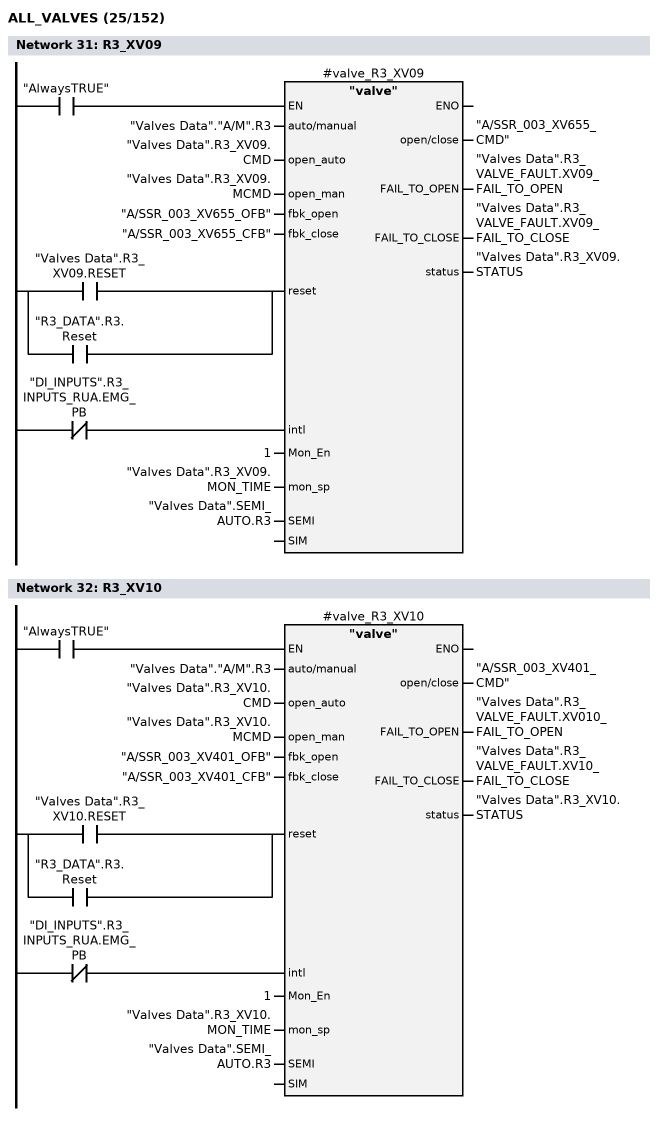
   RUNG wire#powerrail
      Contact( "AlwaysTRUE" )
      #valve_R3_XV09(reset := wire#w1, intl := wire#w2, "auto/manual" := "Valves Data"."A/M".R3, open_auto := "Valves Data".R3_XV09.CMD, open_man := "Valves Data".R3_XV09.MCMD, fbk_open := "A/SSR_003_XV655_OFB", fbk_close := "A/SSR_003_XV655_CFB", Mon_En := 1, mon_sp := "Valves Data".R3_XV09.MON_TIME, SEMI := "Valves Data".SEMI_AUTO.R3, SIM :=, "open/close" => "A/SSR_003_XV655_CMD", FAIL_TO_OPEN => "Valves Data".R3_VALVE_FAULT.XV09_FAIL_TO_OPEN, FAIL_TO_CLOSE => "Valves Data".R3_VALVE_FAULT.XV09_FAIL_TO_CLOSE, status => "Valves Data".R3_XV09.STATUS)
   END_RUNG
   RUNG wire#powerrail
      Contact( "Valves Data".R3_XV09.RESET )
   END_RUNG wire#w1
   RUNG wire#powerrail
      Contact( "R3_DATA".R3.Reset )
   END_RUNG wire#w1
   RUNG wire#powerrail
      I_Contact( "DI_INPUTS".R3_INPUTS_RUA.EMG_PB )
   END_RUNG wire#w2
   // the same network as SCL:
   IF "AlwaysTRUE" THEN
       #valve_R3_XV09("auto/manual" := "Valves Data"."A/M".R3,   // "valve"
                      open_auto := "Valves Data".R3_XV09.CMD,
                      open_man := "Valves Data".R3_XV09.MCMD,
                      fbk_open := "A/SSR_003_XV655_OFB",
                      fbk_close := "A/SSR_003_XV655_CFB",
                      reset := "Valves Data".R3_XV09.RESET OR "R3_DATA".R3.Reset,
                      intl := NOT "DI_INPUTS".R3_INPUTS_RUA.EMG_PB,
                      Mon_En := 1,
                      mon_sp := "Valves Data".R3_XV09.MON_TIME,
                      SEMI := "Valves Data".SEMI_AUTO.R3,
                      "open/close" => "A/SSR_003_XV655_CMD",
                      FAIL_TO_OPEN => "Valves Data".R3_VALVE_FAULT.XV09_FAIL_TO_OPEN,
                      FAIL_TO_CLOSE => "Valves Data".R3_VALVE_FAULT.XV09_FAIL_TO_CLOSE,
                      status => "Valves Data".R3_XV09.STATUS);
   END_IF;
END_REGION

REGION Network 32: R3_XV10
   RUNG wire#powerrail
      Contact( "AlwaysTRUE" )
      #valve_R3_XV10(reset := wire#w1, intl := wire#w2, "auto/manual" := "Valves Data"."A/M".R3, open_auto := "Valves Data".R3_XV10.CMD, open_man := "Valves Data".R3_XV10.MCMD, fbk_open := "A/SSR_003_XV401_OFB", fbk_close := "A/SSR_003_XV401_CFB", Mon_En := 1, mon_sp := "Valves Data".R3_XV10.MON_TIME, SEMI := "Valves Data".SEMI_AUTO.R3, SIM :=, "open/close" => "A/SSR_003_XV401_CMD", FAIL_TO_OPEN => "Valves Data".R3_VALVE_FAULT.XV010_FAIL_TO_OPEN, FAIL_TO_CLOSE => "Valves Data".R3_VALVE_FAULT.XV10_FAIL_TO_CLOSE, status => "Valves Data".R3_XV10.STATUS)
   END_RUNG
   RUNG wire#powerrail
      Contact( "Valves Data".R3_XV10.RESET )
   END_RUNG wire#w1
   RUNG wire#powerrail
      Contact( "R3_DATA".R3.Reset )
   END_RUNG wire#w1
   RUNG wire#powerrail
      I_Contact( "DI_INPUTS".R3_INPUTS_RUA.EMG_PB )
   END_RUNG wire#w2
   // the same network as SCL:
   IF "AlwaysTRUE" THEN
       #valve_R3_XV10("auto/manual" := "Valves Data"."A/M".R3,   // "valve"
                      open_auto := "Valves Data".R3_XV10.CMD,
                      open_man := "Valves Data".R3_XV10.MCMD,
                      fbk_open := "A/SSR_003_XV401_OFB",
                      fbk_close := "A/SSR_003_XV401_CFB",
                      reset := "Valves Data".R3_XV10.RESET OR "R3_DATA".R3.Reset,
                      intl := NOT "DI_INPUTS".R3_INPUTS_RUA.EMG_PB,
                      Mon_En := 1,
                      mon_sp := "Valves Data".R3_XV10.MON_TIME,
                      SEMI := "Valves Data".SEMI_AUTO.R3,
                      "open/close" => "A/SSR_003_XV401_CMD",
                      FAIL_TO_OPEN => "Valves Data".R3_VALVE_FAULT.XV010_FAIL_TO_OPEN,
                      FAIL_TO_CLOSE => "Valves Data".R3_VALVE_FAULT.XV10_FAIL_TO_CLOSE,
                      status => "Valves Data".R3_XV10.STATUS);
   END_IF;
END_REGION

REGION Network 33: ****REACTOR_04****
END_REGION

REGION Network 34: R4_XV01
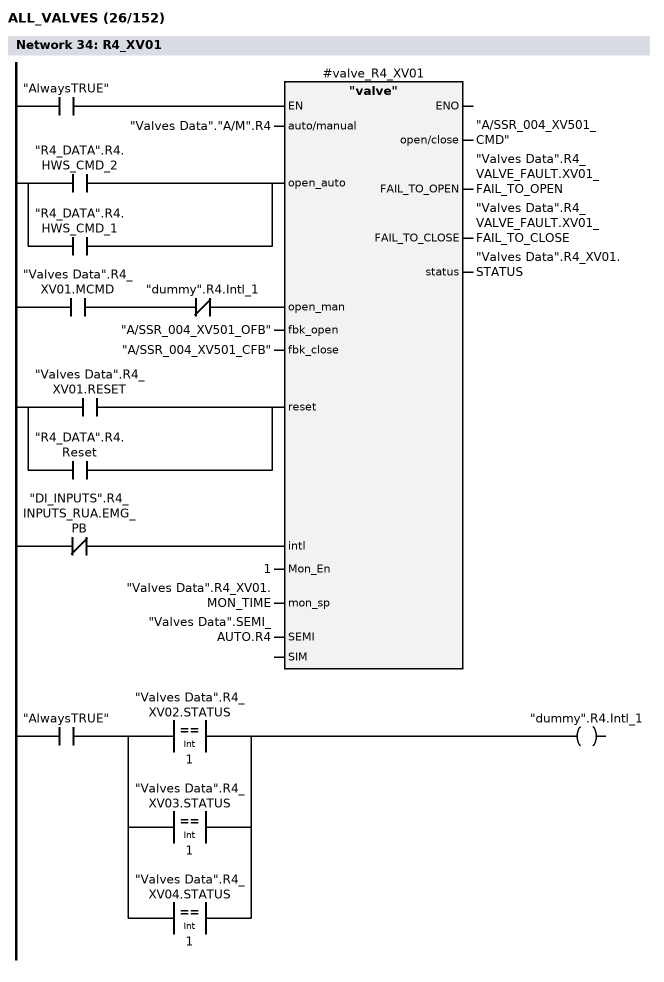
   RUNG wire#powerrail
      Contact( "AlwaysTRUE" )
      #valve_R4_XV01(open_auto := wire#w1, open_man := wire#w2, reset := wire#w3, intl := wire#w4, "auto/manual" := "Valves Data"."A/M".R4, fbk_open := "A/SSR_004_XV501_OFB", fbk_close := "A/SSR_004_XV501_CFB", Mon_En := 1, mon_sp := "Valves Data".R4_XV01.MON_TIME, SEMI := "Valves Data".SEMI_AUTO.R4, SIM :=, "open/close" => "A/SSR_004_XV501_CMD", FAIL_TO_OPEN => "Valves Data".R4_VALVE_FAULT.XV01_FAIL_TO_OPEN, FAIL_TO_CLOSE => "Valves Data".R4_VALVE_FAULT.XV01_FAIL_TO_CLOSE, status => "Valves Data".R4_XV01.STATUS)
   END_RUNG
   RUNG wire#powerrail
      Contact( "R4_DATA".R4.HWS_CMD_2 )
   END_RUNG wire#w1
   RUNG wire#powerrail
      Contact( "R4_DATA".R4.HWS_CMD_1 )
   END_RUNG wire#w1
   RUNG wire#powerrail
      Contact( "Valves Data".R4_XV01.MCMD )
      I_Contact( "dummy".R4.Intl_1 )
   END_RUNG wire#w2
   RUNG wire#powerrail
      Contact( "Valves Data".R4_XV01.RESET )
   END_RUNG wire#w3
   RUNG wire#powerrail
      Contact( "R4_DATA".R4.Reset )
   END_RUNG wire#w3
   RUNG wire#powerrail
      I_Contact( "DI_INPUTS".R4_INPUTS_RUA.EMG_PB )
   END_RUNG wire#w4
   RUNG wire#powerrail
      Contact( "AlwaysTRUE" )
      wire#w5
      { S7_Templates := "SrcType := Int" } EQ_Contact(in1 := "Valves Data".R4_XV02.STATUS, in2 := 1)
      wire#w6
      Coil( "dummy".R4.Intl_1 )
   END_RUNG
   RUNG wire#w5
      { S7_Templates := "SrcType := Int" } EQ_Contact(in1 := "Valves Data".R4_XV03.STATUS, in2 := 1)
   END_RUNG wire#w6
   RUNG wire#w5
      { S7_Templates := "SrcType := Int" } EQ_Contact(in1 := "Valves Data".R4_XV04.STATUS, in2 := 1)
   END_RUNG wire#w6
   // the same network as SCL:
   IF "AlwaysTRUE" THEN
       #valve_R4_XV01("auto/manual" := "Valves Data"."A/M".R4,   // "valve"
                      open_auto := "R4_DATA".R4.HWS_CMD_2 OR "R4_DATA".R4.HWS_CMD_1,
                      open_man := "Valves Data".R4_XV01.MCMD AND NOT "dummy".R4.Intl_1,
                      fbk_open := "A/SSR_004_XV501_OFB",
                      fbk_close := "A/SSR_004_XV501_CFB",
                      reset := "Valves Data".R4_XV01.RESET OR "R4_DATA".R4.Reset,
                      intl := NOT "DI_INPUTS".R4_INPUTS_RUA.EMG_PB,
                      Mon_En := 1,
                      mon_sp := "Valves Data".R4_XV01.MON_TIME,
                      SEMI := "Valves Data".SEMI_AUTO.R4,
                      "open/close" => "A/SSR_004_XV501_CMD",
                      FAIL_TO_OPEN => "Valves Data".R4_VALVE_FAULT.XV01_FAIL_TO_OPEN,
                      FAIL_TO_CLOSE => "Valves Data".R4_VALVE_FAULT.XV01_FAIL_TO_CLOSE,
                      status => "Valves Data".R4_XV01.STATUS);
   END_IF;
   "dummy".R4.Intl_1 := "AlwaysTRUE" AND (("Valves Data".R4_XV02.STATUS = 1) OR ("Valves Data".R4_XV03.STATUS = 1) OR ("Valves Data".R4_XV04.STATUS = 1));
END_REGION

REGION Network 35: R4_XV02
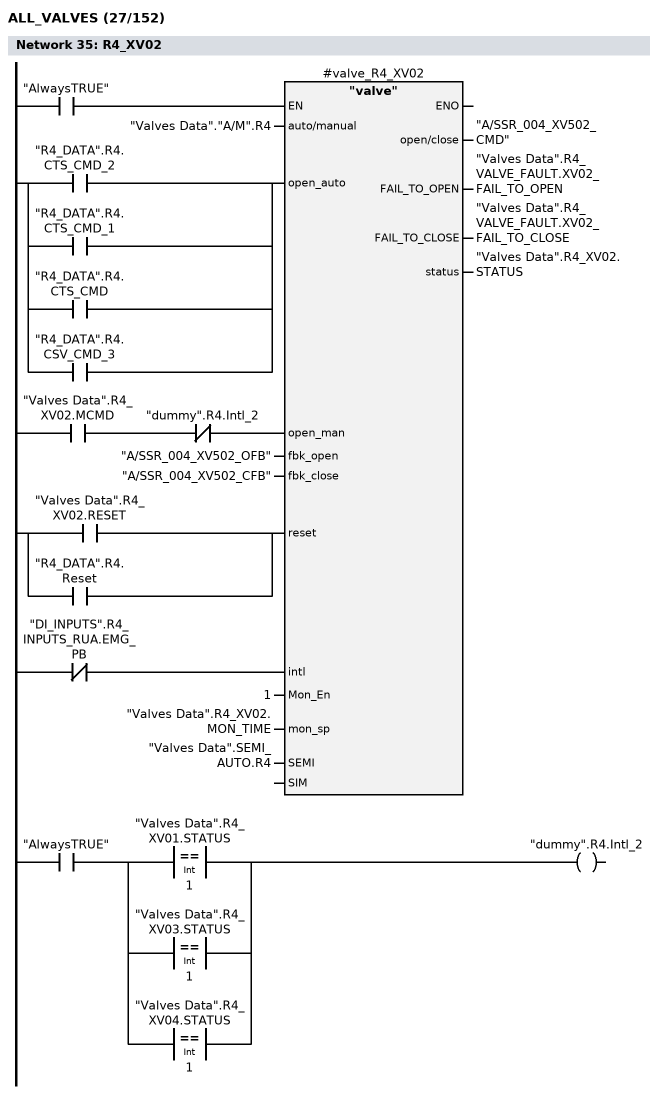
   RUNG wire#powerrail
      Contact( "AlwaysTRUE" )
      #valve_R4_XV02(open_auto := wire#w1, open_man := wire#w2, reset := wire#w3, intl := wire#w4, "auto/manual" := "Valves Data"."A/M".R4, fbk_open := "A/SSR_004_XV502_OFB", fbk_close := "A/SSR_004_XV502_CFB", Mon_En := 1, mon_sp := "Valves Data".R4_XV02.MON_TIME, SEMI := "Valves Data".SEMI_AUTO.R4, SIM :=, "open/close" => "A/SSR_004_XV502_CMD", FAIL_TO_OPEN => "Valves Data".R4_VALVE_FAULT.XV02_FAIL_TO_OPEN, FAIL_TO_CLOSE => "Valves Data".R4_VALVE_FAULT.XV02_FAIL_TO_CLOSE, status => "Valves Data".R4_XV02.STATUS)
   END_RUNG
   RUNG wire#powerrail
      Contact( "R4_DATA".R4.CTS_CMD_2 )
   END_RUNG wire#w1
   RUNG wire#powerrail
      Contact( "R4_DATA".R4.CTS_CMD_1 )
   END_RUNG wire#w1
   RUNG wire#powerrail
      Contact( "R4_DATA".R4.CTS_CMD )
   END_RUNG wire#w1
   RUNG wire#powerrail
      Contact( "R4_DATA".R4.CSV_CMD_3 )
   END_RUNG wire#w1
   RUNG wire#powerrail
      Contact( "Valves Data".R4_XV02.MCMD )
      I_Contact( "dummy".R4.Intl_2 )
   END_RUNG wire#w2
   RUNG wire#powerrail
      Contact( "Valves Data".R4_XV02.RESET )
   END_RUNG wire#w3
   RUNG wire#powerrail
      Contact( "R4_DATA".R4.Reset )
   END_RUNG wire#w3
   RUNG wire#powerrail
      I_Contact( "DI_INPUTS".R4_INPUTS_RUA.EMG_PB )
   END_RUNG wire#w4
   RUNG wire#powerrail
      Contact( "AlwaysTRUE" )
      wire#w5
      { S7_Templates := "SrcType := Int" } EQ_Contact(in1 := "Valves Data".R4_XV01.STATUS, in2 := 1)
      wire#w6
      Coil( "dummy".R4.Intl_2 )
   END_RUNG
   RUNG wire#w5
      { S7_Templates := "SrcType := Int" } EQ_Contact(in1 := "Valves Data".R4_XV03.STATUS, in2 := 1)
   END_RUNG wire#w6
   RUNG wire#w5
      { S7_Templates := "SrcType := Int" } EQ_Contact(in1 := "Valves Data".R4_XV04.STATUS, in2 := 1)
   END_RUNG wire#w6
   // the same network as SCL:
   IF "AlwaysTRUE" THEN
       #valve_R4_XV02("auto/manual" := "Valves Data"."A/M".R4,   // "valve"
                      open_auto := "R4_DATA".R4.CTS_CMD_2 OR "R4_DATA".R4.CTS_CMD_1 OR "R4_DATA".R4.CTS_CMD OR "R4_DATA".R4.CSV_CMD_3,
                      open_man := "Valves Data".R4_XV02.MCMD AND NOT "dummy".R4.Intl_2,
                      fbk_open := "A/SSR_004_XV502_OFB",
                      fbk_close := "A/SSR_004_XV502_CFB",
                      reset := "Valves Data".R4_XV02.RESET OR "R4_DATA".R4.Reset,
                      intl := NOT "DI_INPUTS".R4_INPUTS_RUA.EMG_PB,
                      Mon_En := 1,
                      mon_sp := "Valves Data".R4_XV02.MON_TIME,
                      SEMI := "Valves Data".SEMI_AUTO.R4,
                      "open/close" => "A/SSR_004_XV502_CMD",
                      FAIL_TO_OPEN => "Valves Data".R4_VALVE_FAULT.XV02_FAIL_TO_OPEN,
                      FAIL_TO_CLOSE => "Valves Data".R4_VALVE_FAULT.XV02_FAIL_TO_CLOSE,
                      status => "Valves Data".R4_XV02.STATUS);
   END_IF;
   "dummy".R4.Intl_2 := "AlwaysTRUE" AND (("Valves Data".R4_XV01.STATUS = 1) OR ("Valves Data".R4_XV03.STATUS = 1) OR ("Valves Data".R4_XV04.STATUS = 1));
END_REGION

REGION Network 36: R4_XV03
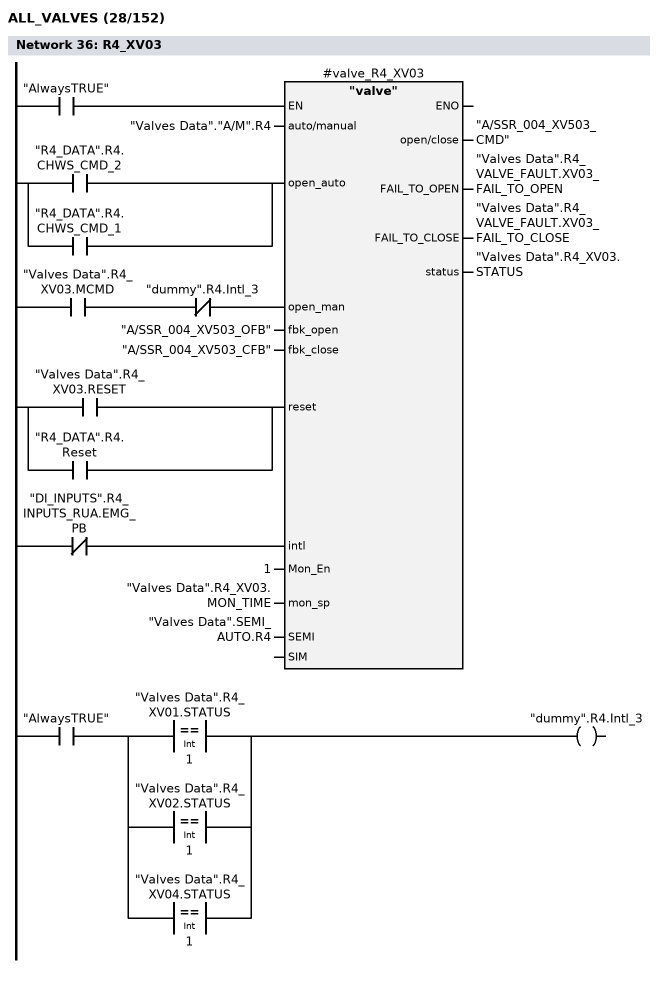
   RUNG wire#powerrail
      Contact( "AlwaysTRUE" )
      #valve_R4_XV03(open_auto := wire#w1, open_man := wire#w2, reset := wire#w3, intl := wire#w4, "auto/manual" := "Valves Data"."A/M".R4, fbk_open := "A/SSR_004_XV503_OFB", fbk_close := "A/SSR_004_XV503_CFB", Mon_En := 1, mon_sp := "Valves Data".R4_XV03.MON_TIME, SEMI := "Valves Data".SEMI_AUTO.R4, SIM :=, "open/close" => "A/SSR_004_XV503_CMD", FAIL_TO_OPEN => "Valves Data".R4_VALVE_FAULT.XV03_FAIL_TO_OPEN, FAIL_TO_CLOSE => "Valves Data".R4_VALVE_FAULT.XV03_FAIL_TO_CLOSE, status => "Valves Data".R4_XV03.STATUS)
   END_RUNG
   RUNG wire#powerrail
      Contact( "R4_DATA".R4.CHWS_CMD_2 )
   END_RUNG wire#w1
   RUNG wire#powerrail
      Contact( "R4_DATA".R4.CHWS_CMD_1 )
   END_RUNG wire#w1
   RUNG wire#powerrail
      Contact( "Valves Data".R4_XV03.MCMD )
      I_Contact( "dummy".R4.Intl_3 )
   END_RUNG wire#w2
   RUNG wire#powerrail
      Contact( "Valves Data".R4_XV03.RESET )
   END_RUNG wire#w3
   RUNG wire#powerrail
      Contact( "R4_DATA".R4.Reset )
   END_RUNG wire#w3
   RUNG wire#powerrail
      I_Contact( "DI_INPUTS".R4_INPUTS_RUA.EMG_PB )
   END_RUNG wire#w4
   RUNG wire#powerrail
      Contact( "AlwaysTRUE" )
      wire#w5
      { S7_Templates := "SrcType := Int" } EQ_Contact(in1 := "Valves Data".R4_XV01.STATUS, in2 := 1)
      wire#w6
      Coil( "dummy".R4.Intl_3 )
   END_RUNG
   RUNG wire#w5
      { S7_Templates := "SrcType := Int" } EQ_Contact(in1 := "Valves Data".R4_XV02.STATUS, in2 := 1)
   END_RUNG wire#w6
   RUNG wire#w5
      { S7_Templates := "SrcType := Int" } EQ_Contact(in1 := "Valves Data".R4_XV04.STATUS, in2 := 1)
   END_RUNG wire#w6
   // the same network as SCL:
   IF "AlwaysTRUE" THEN
       #valve_R4_XV03("auto/manual" := "Valves Data"."A/M".R4,   // "valve"
                      open_auto := "R4_DATA".R4.CHWS_CMD_2 OR "R4_DATA".R4.CHWS_CMD_1,
                      open_man := "Valves Data".R4_XV03.MCMD AND NOT "dummy".R4.Intl_3,
                      fbk_open := "A/SSR_004_XV503_OFB",
                      fbk_close := "A/SSR_004_XV503_CFB",
                      reset := "Valves Data".R4_XV03.RESET OR "R4_DATA".R4.Reset,
                      intl := NOT "DI_INPUTS".R4_INPUTS_RUA.EMG_PB,
                      Mon_En := 1,
                      mon_sp := "Valves Data".R4_XV03.MON_TIME,
                      SEMI := "Valves Data".SEMI_AUTO.R4,
                      "open/close" => "A/SSR_004_XV503_CMD",
                      FAIL_TO_OPEN => "Valves Data".R4_VALVE_FAULT.XV03_FAIL_TO_OPEN,
                      FAIL_TO_CLOSE => "Valves Data".R4_VALVE_FAULT.XV03_FAIL_TO_CLOSE,
                      status => "Valves Data".R4_XV03.STATUS);
   END_IF;
   "dummy".R4.Intl_3 := "AlwaysTRUE" AND (("Valves Data".R4_XV01.STATUS = 1) OR ("Valves Data".R4_XV02.STATUS = 1) OR ("Valves Data".R4_XV04.STATUS = 1));
END_REGION

REGION Network 37: R4_XV04
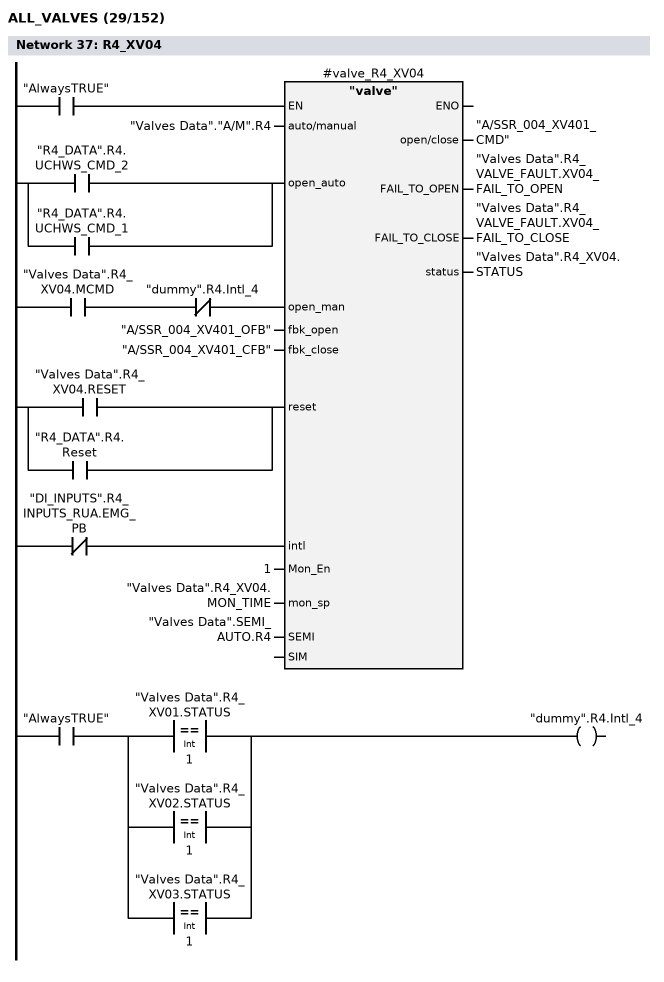
   RUNG wire#powerrail
      Contact( "AlwaysTRUE" )
      #valve_R4_XV04(open_auto := wire#w1, open_man := wire#w2, reset := wire#w3, intl := wire#w4, "auto/manual" := "Valves Data"."A/M".R4, fbk_open := "A/SSR_004_XV401_OFB", fbk_close := "A/SSR_004_XV401_CFB", Mon_En := 1, mon_sp := "Valves Data".R4_XV04.MON_TIME, SEMI := "Valves Data".SEMI_AUTO.R4, SIM :=, "open/close" => "A/SSR_004_XV401_CMD", FAIL_TO_OPEN => "Valves Data".R4_VALVE_FAULT.XV04_FAIL_TO_OPEN, FAIL_TO_CLOSE => "Valves Data".R4_VALVE_FAULT.XV04_FAIL_TO_CLOSE, status => "Valves Data".R4_XV04.STATUS)
   END_RUNG
   RUNG wire#powerrail
      Contact( "R4_DATA".R4.UCHWS_CMD_2 )
   END_RUNG wire#w1
   RUNG wire#powerrail
      Contact( "R4_DATA".R4.UCHWS_CMD_1 )
   END_RUNG wire#w1
   RUNG wire#powerrail
      Contact( "Valves Data".R4_XV04.MCMD )
      I_Contact( "dummy".R4.Intl_4 )
   END_RUNG wire#w2
   RUNG wire#powerrail
      Contact( "Valves Data".R4_XV04.RESET )
   END_RUNG wire#w3
   RUNG wire#powerrail
      Contact( "R4_DATA".R4.Reset )
   END_RUNG wire#w3
   RUNG wire#powerrail
      I_Contact( "DI_INPUTS".R4_INPUTS_RUA.EMG_PB )
   END_RUNG wire#w4
   RUNG wire#powerrail
      Contact( "AlwaysTRUE" )
      wire#w5
      { S7_Templates := "SrcType := Int" } EQ_Contact(in1 := "Valves Data".R4_XV01.STATUS, in2 := 1)
      wire#w6
      Coil( "dummy".R4.Intl_4 )
   END_RUNG
   RUNG wire#w5
      { S7_Templates := "SrcType := Int" } EQ_Contact(in1 := "Valves Data".R4_XV02.STATUS, in2 := 1)
   END_RUNG wire#w6
   RUNG wire#w5
      { S7_Templates := "SrcType := Int" } EQ_Contact(in1 := "Valves Data".R4_XV03.STATUS, in2 := 1)
   END_RUNG wire#w6
   // the same network as SCL:
   IF "AlwaysTRUE" THEN
       #valve_R4_XV04("auto/manual" := "Valves Data"."A/M".R4,   // "valve"
                      open_auto := "R4_DATA".R4.UCHWS_CMD_2 OR "R4_DATA".R4.UCHWS_CMD_1,
                      open_man := "Valves Data".R4_XV04.MCMD AND NOT "dummy".R4.Intl_4,
                      fbk_open := "A/SSR_004_XV401_OFB",
                      fbk_close := "A/SSR_004_XV401_CFB",
                      reset := "Valves Data".R4_XV04.RESET OR "R4_DATA".R4.Reset,
                      intl := NOT "DI_INPUTS".R4_INPUTS_RUA.EMG_PB,
                      Mon_En := 1,
                      mon_sp := "Valves Data".R4_XV04.MON_TIME,
                      SEMI := "Valves Data".SEMI_AUTO.R4,
                      "open/close" => "A/SSR_004_XV401_CMD",
                      FAIL_TO_OPEN => "Valves Data".R4_VALVE_FAULT.XV04_FAIL_TO_OPEN,
                      FAIL_TO_CLOSE => "Valves Data".R4_VALVE_FAULT.XV04_FAIL_TO_CLOSE,
                      status => "Valves Data".R4_XV04.STATUS);
   END_IF;
   "dummy".R4.Intl_4 := "AlwaysTRUE" AND (("Valves Data".R4_XV01.STATUS = 1) OR ("Valves Data".R4_XV02.STATUS = 1) OR ("Valves Data".R4_XV03.STATUS = 1));
END_REGION

REGION Network 38: R4_XV05
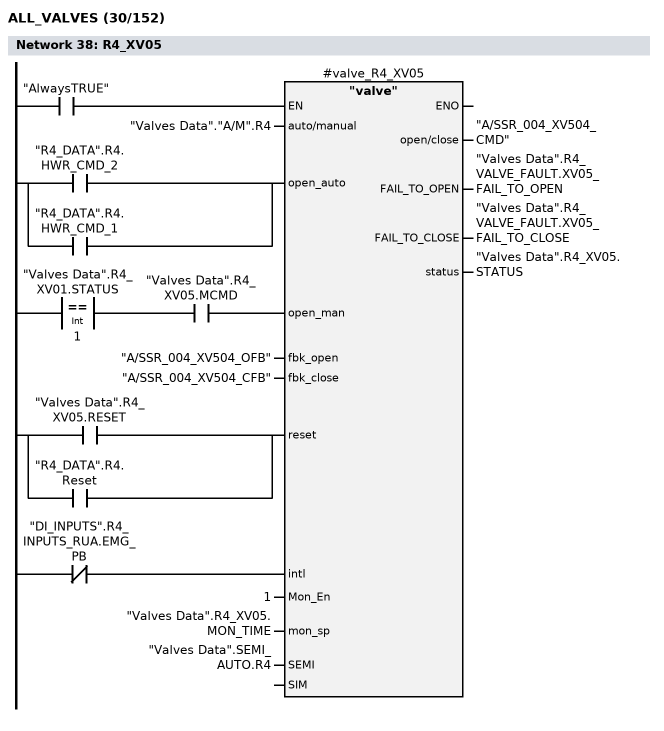
   RUNG wire#powerrail
      Contact( "AlwaysTRUE" )
      #valve_R4_XV05(open_auto := wire#w1, open_man := wire#w2, reset := wire#w3, intl := wire#w4, "auto/manual" := "Valves Data"."A/M".R4, fbk_open := "A/SSR_004_XV504_OFB", fbk_close := "A/SSR_004_XV504_CFB", Mon_En := 1, mon_sp := "Valves Data".R4_XV05.MON_TIME, SEMI := "Valves Data".SEMI_AUTO.R4, SIM :=, "open/close" => "A/SSR_004_XV504_CMD", FAIL_TO_OPEN => "Valves Data".R4_VALVE_FAULT.XV05_FAIL_TO_OPEN, FAIL_TO_CLOSE => "Valves Data".R4_VALVE_FAULT.XV05_FAIL_TO_CLOSE, status => "Valves Data".R4_XV05.STATUS)
   END_RUNG
   RUNG wire#powerrail
      Contact( "R4_DATA".R4.HWR_CMD_2 )
   END_RUNG wire#w1
   RUNG wire#powerrail
      Contact( "R4_DATA".R4.HWR_CMD_1 )
   END_RUNG wire#w1
   RUNG wire#powerrail
      { S7_Templates := "SrcType := Int" } EQ_Contact(in1 := "Valves Data".R4_XV01.STATUS, in2 := 1)
      Contact( "Valves Data".R4_XV05.MCMD )
   END_RUNG wire#w2
   RUNG wire#powerrail
      Contact( "Valves Data".R4_XV05.RESET )
   END_RUNG wire#w3
   RUNG wire#powerrail
      Contact( "R4_DATA".R4.Reset )
   END_RUNG wire#w3
   RUNG wire#powerrail
      I_Contact( "DI_INPUTS".R4_INPUTS_RUA.EMG_PB )
   END_RUNG wire#w4
   // the same network as SCL:
   IF "AlwaysTRUE" THEN
       #valve_R4_XV05("auto/manual" := "Valves Data"."A/M".R4,   // "valve"
                      open_auto := "R4_DATA".R4.HWR_CMD_2 OR "R4_DATA".R4.HWR_CMD_1,
                      open_man := ("Valves Data".R4_XV01.STATUS = 1) AND "Valves Data".R4_XV05.MCMD,
                      fbk_open := "A/SSR_004_XV504_OFB",
                      fbk_close := "A/SSR_004_XV504_CFB",
                      reset := "Valves Data".R4_XV05.RESET OR "R4_DATA".R4.Reset,
                      intl := NOT "DI_INPUTS".R4_INPUTS_RUA.EMG_PB,
                      Mon_En := 1,
                      mon_sp := "Valves Data".R4_XV05.MON_TIME,
                      SEMI := "Valves Data".SEMI_AUTO.R4,
                      "open/close" => "A/SSR_004_XV504_CMD",
                      FAIL_TO_OPEN => "Valves Data".R4_VALVE_FAULT.XV05_FAIL_TO_OPEN,
                      FAIL_TO_CLOSE => "Valves Data".R4_VALVE_FAULT.XV05_FAIL_TO_CLOSE,
                      status => "Valves Data".R4_XV05.STATUS);
   END_IF;
END_REGION

REGION Network 39: R4_XV06
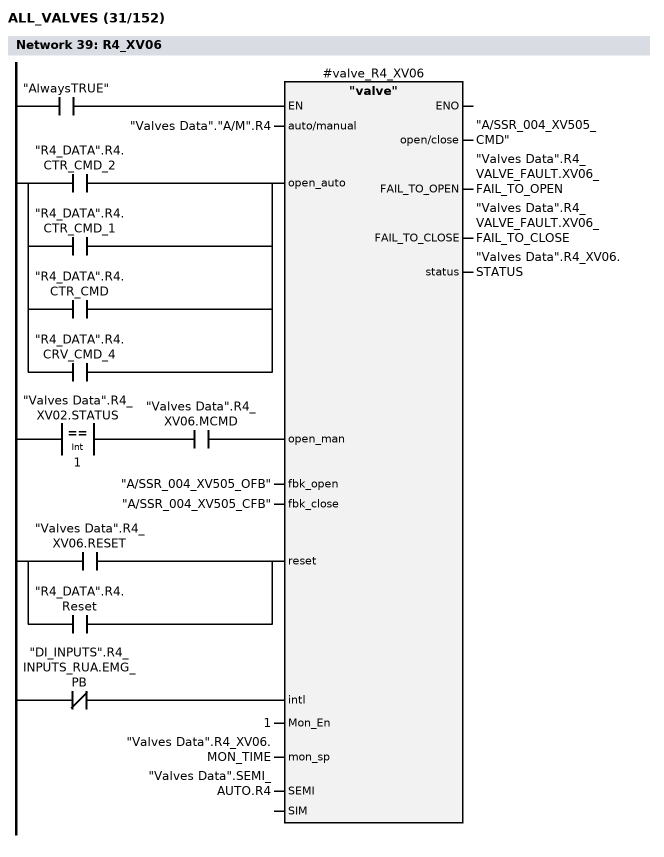
   RUNG wire#powerrail
      Contact( "AlwaysTRUE" )
      #valve_R4_XV06(open_auto := wire#w1, open_man := wire#w2, reset := wire#w3, intl := wire#w4, "auto/manual" := "Valves Data"."A/M".R4, fbk_open := "A/SSR_004_XV505_OFB", fbk_close := "A/SSR_004_XV505_CFB", Mon_En := 1, mon_sp := "Valves Data".R4_XV06.MON_TIME, SEMI := "Valves Data".SEMI_AUTO.R4, SIM :=, "open/close" => "A/SSR_004_XV505_CMD", FAIL_TO_OPEN => "Valves Data".R4_VALVE_FAULT.XV06_FAIL_TO_OPEN, FAIL_TO_CLOSE => "Valves Data".R4_VALVE_FAULT.XV06_FAIL_TO_CLOSE, status => "Valves Data".R4_XV06.STATUS)
   END_RUNG
   RUNG wire#powerrail
      Contact( "R4_DATA".R4.CTR_CMD_2 )
   END_RUNG wire#w1
   RUNG wire#powerrail
      Contact( "R4_DATA".R4.CTR_CMD_1 )
   END_RUNG wire#w1
   RUNG wire#powerrail
      Contact( "R4_DATA".R4.CTR_CMD )
   END_RUNG wire#w1
   RUNG wire#powerrail
      Contact( "R4_DATA".R4.CRV_CMD_4 )
   END_RUNG wire#w1
   RUNG wire#powerrail
      { S7_Templates := "SrcType := Int" } EQ_Contact(in1 := "Valves Data".R4_XV02.STATUS, in2 := 1)
      Contact( "Valves Data".R4_XV06.MCMD )
   END_RUNG wire#w2
   RUNG wire#powerrail
      Contact( "Valves Data".R4_XV06.RESET )
   END_RUNG wire#w3
   RUNG wire#powerrail
      Contact( "R4_DATA".R4.Reset )
   END_RUNG wire#w3
   RUNG wire#powerrail
      I_Contact( "DI_INPUTS".R4_INPUTS_RUA.EMG_PB )
   END_RUNG wire#w4
   // the same network as SCL:
   IF "AlwaysTRUE" THEN
       #valve_R4_XV06("auto/manual" := "Valves Data"."A/M".R4,   // "valve"
                      open_auto := "R4_DATA".R4.CTR_CMD_2 OR "R4_DATA".R4.CTR_CMD_1 OR "R4_DATA".R4.CTR_CMD OR "R4_DATA".R4.CRV_CMD_4,
                      open_man := ("Valves Data".R4_XV02.STATUS = 1) AND "Valves Data".R4_XV06.MCMD,
                      fbk_open := "A/SSR_004_XV505_OFB",
                      fbk_close := "A/SSR_004_XV505_CFB",
                      reset := "Valves Data".R4_XV06.RESET OR "R4_DATA".R4.Reset,
                      intl := NOT "DI_INPUTS".R4_INPUTS_RUA.EMG_PB,
                      Mon_En := 1,
                      mon_sp := "Valves Data".R4_XV06.MON_TIME,
                      SEMI := "Valves Data".SEMI_AUTO.R4,
                      "open/close" => "A/SSR_004_XV505_CMD",
                      FAIL_TO_OPEN => "Valves Data".R4_VALVE_FAULT.XV06_FAIL_TO_OPEN,
                      FAIL_TO_CLOSE => "Valves Data".R4_VALVE_FAULT.XV06_FAIL_TO_CLOSE,
                      status => "Valves Data".R4_XV06.STATUS);
   END_IF;
END_REGION

REGION Network 40: R4_XV07
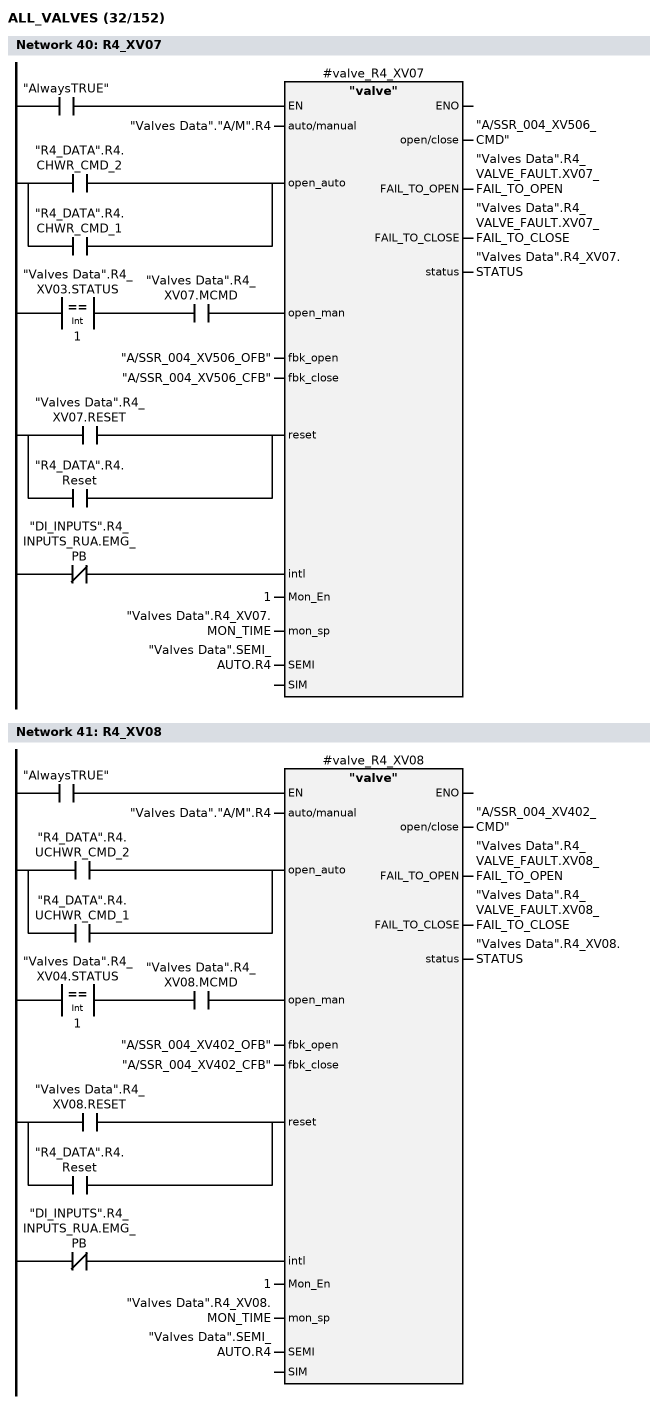
   RUNG wire#powerrail
      Contact( "AlwaysTRUE" )
      #valve_R4_XV07(open_auto := wire#w1, open_man := wire#w2, reset := wire#w3, intl := wire#w4, "auto/manual" := "Valves Data"."A/M".R4, fbk_open := "A/SSR_004_XV506_OFB", fbk_close := "A/SSR_004_XV506_CFB", Mon_En := 1, mon_sp := "Valves Data".R4_XV07.MON_TIME, SEMI := "Valves Data".SEMI_AUTO.R4, SIM :=, "open/close" => "A/SSR_004_XV506_CMD", FAIL_TO_OPEN => "Valves Data".R4_VALVE_FAULT.XV07_FAIL_TO_OPEN, FAIL_TO_CLOSE => "Valves Data".R4_VALVE_FAULT.XV07_FAIL_TO_CLOSE, status => "Valves Data".R4_XV07.STATUS)
   END_RUNG
   RUNG wire#powerrail
      Contact( "R4_DATA".R4.CHWR_CMD_2 )
   END_RUNG wire#w1
   RUNG wire#powerrail
      Contact( "R4_DATA".R4.CHWR_CMD_1 )
   END_RUNG wire#w1
   RUNG wire#powerrail
      { S7_Templates := "SrcType := Int" } EQ_Contact(in1 := "Valves Data".R4_XV03.STATUS, in2 := 1)
      Contact( "Valves Data".R4_XV07.MCMD )
   END_RUNG wire#w2
   RUNG wire#powerrail
      Contact( "Valves Data".R4_XV07.RESET )
   END_RUNG wire#w3
   RUNG wire#powerrail
      Contact( "R4_DATA".R4.Reset )
   END_RUNG wire#w3
   RUNG wire#powerrail
      I_Contact( "DI_INPUTS".R4_INPUTS_RUA.EMG_PB )
   END_RUNG wire#w4
   // the same network as SCL:
   IF "AlwaysTRUE" THEN
       #valve_R4_XV07("auto/manual" := "Valves Data"."A/M".R4,   // "valve"
                      open_auto := "R4_DATA".R4.CHWR_CMD_2 OR "R4_DATA".R4.CHWR_CMD_1,
                      open_man := ("Valves Data".R4_XV03.STATUS = 1) AND "Valves Data".R4_XV07.MCMD,
                      fbk_open := "A/SSR_004_XV506_OFB",
                      fbk_close := "A/SSR_004_XV506_CFB",
                      reset := "Valves Data".R4_XV07.RESET OR "R4_DATA".R4.Reset,
                      intl := NOT "DI_INPUTS".R4_INPUTS_RUA.EMG_PB,
                      Mon_En := 1,
                      mon_sp := "Valves Data".R4_XV07.MON_TIME,
                      SEMI := "Valves Data".SEMI_AUTO.R4,
                      "open/close" => "A/SSR_004_XV506_CMD",
                      FAIL_TO_OPEN => "Valves Data".R4_VALVE_FAULT.XV07_FAIL_TO_OPEN,
                      FAIL_TO_CLOSE => "Valves Data".R4_VALVE_FAULT.XV07_FAIL_TO_CLOSE,
                      status => "Valves Data".R4_XV07.STATUS);
   END_IF;
END_REGION

REGION Network 41: R4_XV08
   RUNG wire#powerrail
      Contact( "AlwaysTRUE" )
      #valve_R4_XV08(open_auto := wire#w1, open_man := wire#w2, reset := wire#w3, intl := wire#w4, "auto/manual" := "Valves Data"."A/M".R4, fbk_open := "A/SSR_004_XV402_OFB", fbk_close := "A/SSR_004_XV402_CFB", Mon_En := 1, mon_sp := "Valves Data".R4_XV08.MON_TIME, SEMI := "Valves Data".SEMI_AUTO.R4, SIM :=, "open/close" => "A/SSR_004_XV402_CMD", FAIL_TO_OPEN => "Valves Data".R4_VALVE_FAULT.XV08_FAIL_TO_OPEN, FAIL_TO_CLOSE => "Valves Data".R4_VALVE_FAULT.XV08_FAIL_TO_CLOSE, status => "Valves Data".R4_XV08.STATUS)
   END_RUNG
   RUNG wire#powerrail
      Contact( "R4_DATA".R4.UCHWR_CMD_2 )
   END_RUNG wire#w1
   RUNG wire#powerrail
      Contact( "R4_DATA".R4.UCHWR_CMD_1 )
   END_RUNG wire#w1
   RUNG wire#powerrail
      { S7_Templates := "SrcType := Int" } EQ_Contact(in1 := "Valves Data".R4_XV04.STATUS, in2 := 1)
      Contact( "Valves Data".R4_XV08.MCMD )
   END_RUNG wire#w2
   RUNG wire#powerrail
      Contact( "Valves Data".R4_XV08.RESET )
   END_RUNG wire#w3
   RUNG wire#powerrail
      Contact( "R4_DATA".R4.Reset )
   END_RUNG wire#w3
   RUNG wire#powerrail
      I_Contact( "DI_INPUTS".R4_INPUTS_RUA.EMG_PB )
   END_RUNG wire#w4
   // the same network as SCL:
   IF "AlwaysTRUE" THEN
       #valve_R4_XV08("auto/manual" := "Valves Data"."A/M".R4,   // "valve"
                      open_auto := "R4_DATA".R4.UCHWR_CMD_2 OR "R4_DATA".R4.UCHWR_CMD_1,
                      open_man := ("Valves Data".R4_XV04.STATUS = 1) AND "Valves Data".R4_XV08.MCMD,
                      fbk_open := "A/SSR_004_XV402_OFB",
                      fbk_close := "A/SSR_004_XV402_CFB",
                      reset := "Valves Data".R4_XV08.RESET OR "R4_DATA".R4.Reset,
                      intl := NOT "DI_INPUTS".R4_INPUTS_RUA.EMG_PB,
                      Mon_En := 1,
                      mon_sp := "Valves Data".R4_XV08.MON_TIME,
                      SEMI := "Valves Data".SEMI_AUTO.R4,
                      "open/close" => "A/SSR_004_XV402_CMD",
                      FAIL_TO_OPEN => "Valves Data".R4_VALVE_FAULT.XV08_FAIL_TO_OPEN,
                      FAIL_TO_CLOSE => "Valves Data".R4_VALVE_FAULT.XV08_FAIL_TO_CLOSE,
                      status => "Valves Data".R4_XV08.STATUS);
   END_IF;
END_REGION

REGION Network 42: R4_XV09
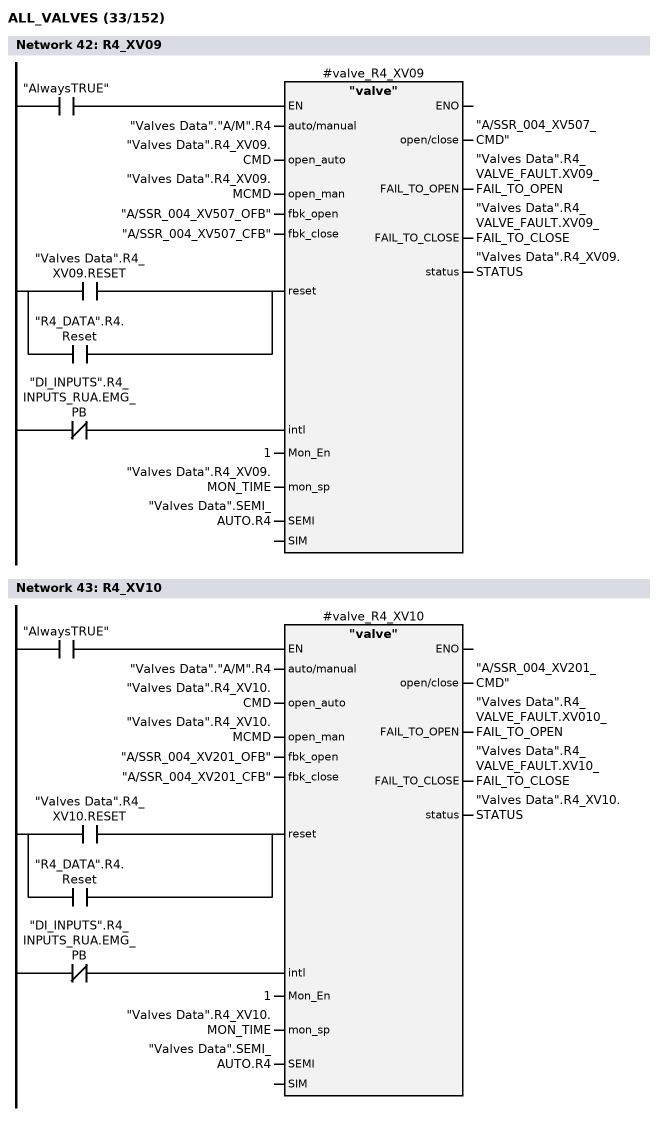
   RUNG wire#powerrail
      Contact( "AlwaysTRUE" )
      #valve_R4_XV09(reset := wire#w1, intl := wire#w2, "auto/manual" := "Valves Data"."A/M".R4, open_auto := "Valves Data".R4_XV09.CMD, open_man := "Valves Data".R4_XV09.MCMD, fbk_open := "A/SSR_004_XV507_OFB", fbk_close := "A/SSR_004_XV507_CFB", Mon_En := 1, mon_sp := "Valves Data".R4_XV09.MON_TIME, SEMI := "Valves Data".SEMI_AUTO.R4, SIM :=, "open/close" => "A/SSR_004_XV507_CMD", FAIL_TO_OPEN => "Valves Data".R4_VALVE_FAULT.XV09_FAIL_TO_OPEN, FAIL_TO_CLOSE => "Valves Data".R4_VALVE_FAULT.XV09_FAIL_TO_CLOSE, status => "Valves Data".R4_XV09.STATUS)
   END_RUNG
   RUNG wire#powerrail
      Contact( "Valves Data".R4_XV09.RESET )
   END_RUNG wire#w1
   RUNG wire#powerrail
      Contact( "R4_DATA".R4.Reset )
   END_RUNG wire#w1
   RUNG wire#powerrail
      I_Contact( "DI_INPUTS".R4_INPUTS_RUA.EMG_PB )
   END_RUNG wire#w2
   // the same network as SCL:
   IF "AlwaysTRUE" THEN
       #valve_R4_XV09("auto/manual" := "Valves Data"."A/M".R4,   // "valve"
                      open_auto := "Valves Data".R4_XV09.CMD,
                      open_man := "Valves Data".R4_XV09.MCMD,
                      fbk_open := "A/SSR_004_XV507_OFB",
                      fbk_close := "A/SSR_004_XV507_CFB",
                      reset := "Valves Data".R4_XV09.RESET OR "R4_DATA".R4.Reset,
                      intl := NOT "DI_INPUTS".R4_INPUTS_RUA.EMG_PB,
                      Mon_En := 1,
                      mon_sp := "Valves Data".R4_XV09.MON_TIME,
                      SEMI := "Valves Data".SEMI_AUTO.R4,
                      "open/close" => "A/SSR_004_XV507_CMD",
                      FAIL_TO_OPEN => "Valves Data".R4_VALVE_FAULT.XV09_FAIL_TO_OPEN,
                      FAIL_TO_CLOSE => "Valves Data".R4_VALVE_FAULT.XV09_FAIL_TO_CLOSE,
                      status => "Valves Data".R4_XV09.STATUS);
   END_IF;
END_REGION

REGION Network 43: R4_XV10
   RUNG wire#powerrail
      Contact( "AlwaysTRUE" )
      #valve_R4_XV10(reset := wire#w1, intl := wire#w2, "auto/manual" := "Valves Data"."A/M".R4, open_auto := "Valves Data".R4_XV10.CMD, open_man := "Valves Data".R4_XV10.MCMD, fbk_open := "A/SSR_004_XV201_OFB", fbk_close := "A/SSR_004_XV201_CFB", Mon_En := 1, mon_sp := "Valves Data".R4_XV10.MON_TIME, SEMI := "Valves Data".SEMI_AUTO.R4, SIM :=, "open/close" => "A/SSR_004_XV201_CMD", FAIL_TO_OPEN => "Valves Data".R4_VALVE_FAULT.XV010_FAIL_TO_OPEN, FAIL_TO_CLOSE => "Valves Data".R4_VALVE_FAULT.XV10_FAIL_TO_CLOSE, status => "Valves Data".R4_XV10.STATUS)
   END_RUNG
   RUNG wire#powerrail
      Contact( "Valves Data".R4_XV10.RESET )
   END_RUNG wire#w1
   RUNG wire#powerrail
      Contact( "R4_DATA".R4.Reset )
   END_RUNG wire#w1
   RUNG wire#powerrail
      I_Contact( "DI_INPUTS".R4_INPUTS_RUA.EMG_PB )
   END_RUNG wire#w2
   // the same network as SCL:
   IF "AlwaysTRUE" THEN
       #valve_R4_XV10("auto/manual" := "Valves Data"."A/M".R4,   // "valve"
                      open_auto := "Valves Data".R4_XV10.CMD,
                      open_man := "Valves Data".R4_XV10.MCMD,
                      fbk_open := "A/SSR_004_XV201_OFB",
                      fbk_close := "A/SSR_004_XV201_CFB",
                      reset := "Valves Data".R4_XV10.RESET OR "R4_DATA".R4.Reset,
                      intl := NOT "DI_INPUTS".R4_INPUTS_RUA.EMG_PB,
                      Mon_En := 1,
                      mon_sp := "Valves Data".R4_XV10.MON_TIME,
                      SEMI := "Valves Data".SEMI_AUTO.R4,
                      "open/close" => "A/SSR_004_XV201_CMD",
                      FAIL_TO_OPEN => "Valves Data".R4_VALVE_FAULT.XV010_FAIL_TO_OPEN,
                      FAIL_TO_CLOSE => "Valves Data".R4_VALVE_FAULT.XV10_FAIL_TO_CLOSE,
                      status => "Valves Data".R4_XV10.STATUS);
   END_IF;
END_REGION

REGION Network 44: ****REACTOR_05****
END_REGION

REGION Network 45: R5_XV01
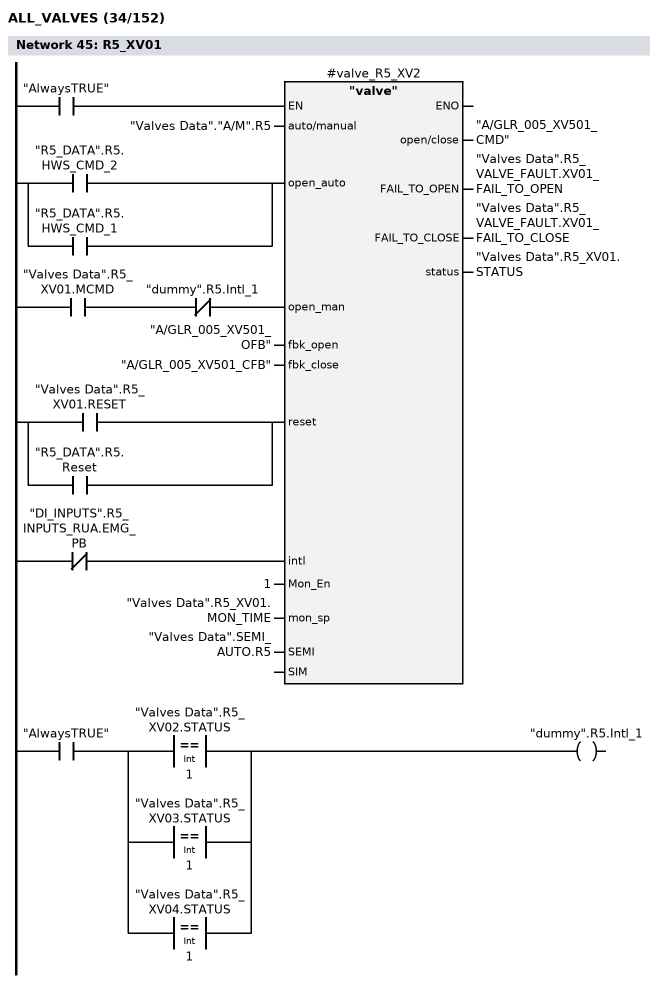
   RUNG wire#powerrail
      Contact( "AlwaysTRUE" )
      #valve_R5_XV2(open_auto := wire#w1, open_man := wire#w2, reset := wire#w3, intl := wire#w4, "auto/manual" := "Valves Data"."A/M".R5, fbk_open := "A/GLR_005_XV501_OFB", fbk_close := "A/GLR_005_XV501_CFB", Mon_En := 1, mon_sp := "Valves Data".R5_XV01.MON_TIME, SEMI := "Valves Data".SEMI_AUTO.R5, SIM :=, "open/close" => "A/GLR_005_XV501_CMD", FAIL_TO_OPEN => "Valves Data".R5_VALVE_FAULT.XV01_FAIL_TO_OPEN, FAIL_TO_CLOSE => "Valves Data".R5_VALVE_FAULT.XV01_FAIL_TO_CLOSE, status => "Valves Data".R5_XV01.STATUS)
   END_RUNG
   RUNG wire#powerrail
      Contact( "R5_DATA".R5.HWS_CMD_2 )
   END_RUNG wire#w1
   RUNG wire#powerrail
      Contact( "R5_DATA".R5.HWS_CMD_1 )
   END_RUNG wire#w1
   RUNG wire#powerrail
      Contact( "Valves Data".R5_XV01.MCMD )
      I_Contact( "dummy".R5.Intl_1 )
   END_RUNG wire#w2
   RUNG wire#powerrail
      Contact( "Valves Data".R5_XV01.RESET )
   END_RUNG wire#w3
   RUNG wire#powerrail
      Contact( "R5_DATA".R5.Reset )
   END_RUNG wire#w3
   RUNG wire#powerrail
      I_Contact( "DI_INPUTS".R5_INPUTS_RUA.EMG_PB )
   END_RUNG wire#w4
   RUNG wire#powerrail
      Contact( "AlwaysTRUE" )
      wire#w5
      { S7_Templates := "SrcType := Int" } EQ_Contact(in1 := "Valves Data".R5_XV02.STATUS, in2 := 1)
      wire#w6
      Coil( "dummy".R5.Intl_1 )
   END_RUNG
   RUNG wire#w5
      { S7_Templates := "SrcType := Int" } EQ_Contact(in1 := "Valves Data".R5_XV03.STATUS, in2 := 1)
   END_RUNG wire#w6
   RUNG wire#w5
      { S7_Templates := "SrcType := Int" } EQ_Contact(in1 := "Valves Data".R5_XV04.STATUS, in2 := 1)
   END_RUNG wire#w6
   // the same network as SCL:
   IF "AlwaysTRUE" THEN
       #valve_R5_XV2("auto/manual" := "Valves Data"."A/M".R5,   // "valve"
                     open_auto := "R5_DATA".R5.HWS_CMD_2 OR "R5_DATA".R5.HWS_CMD_1,
                     open_man := "Valves Data".R5_XV01.MCMD AND NOT "dummy".R5.Intl_1,
                     fbk_open := "A/GLR_005_XV501_OFB",
                     fbk_close := "A/GLR_005_XV501_CFB",
                     reset := "Valves Data".R5_XV01.RESET OR "R5_DATA".R5.Reset,
                     intl := NOT "DI_INPUTS".R5_INPUTS_RUA.EMG_PB,
                     Mon_En := 1,
                     mon_sp := "Valves Data".R5_XV01.MON_TIME,
                     SEMI := "Valves Data".SEMI_AUTO.R5,
                     "open/close" => "A/GLR_005_XV501_CMD",
                     FAIL_TO_OPEN => "Valves Data".R5_VALVE_FAULT.XV01_FAIL_TO_OPEN,
                     FAIL_TO_CLOSE => "Valves Data".R5_VALVE_FAULT.XV01_FAIL_TO_CLOSE,
                     status => "Valves Data".R5_XV01.STATUS);
   END_IF;
   "dummy".R5.Intl_1 := "AlwaysTRUE" AND (("Valves Data".R5_XV02.STATUS = 1) OR ("Valves Data".R5_XV03.STATUS = 1) OR ("Valves Data".R5_XV04.STATUS = 1));
END_REGION

REGION Network 46: R5_XV02
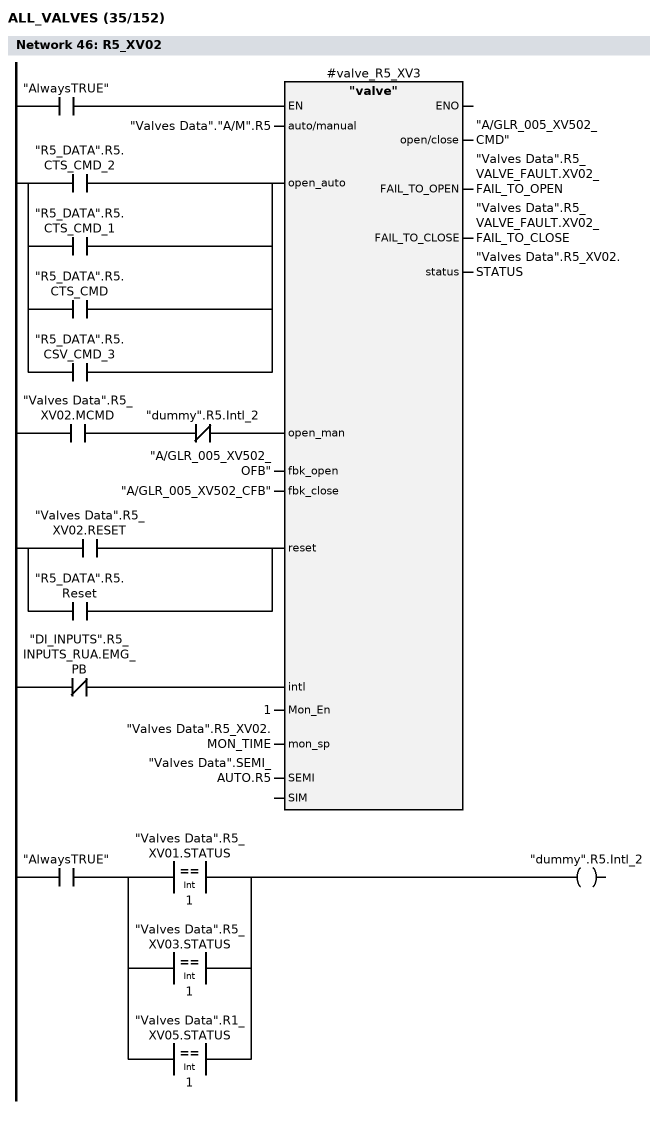
   RUNG wire#powerrail
      Contact( "AlwaysTRUE" )
      #valve_R5_XV3(open_auto := wire#w1, open_man := wire#w2, reset := wire#w3, intl := wire#w4, "auto/manual" := "Valves Data"."A/M".R5, fbk_open := "A/GLR_005_XV502_OFB", fbk_close := "A/GLR_005_XV502_CFB", Mon_En := 1, mon_sp := "Valves Data".R5_XV02.MON_TIME, SEMI := "Valves Data".SEMI_AUTO.R5, SIM :=, "open/close" => "A/GLR_005_XV502_CMD", FAIL_TO_OPEN => "Valves Data".R5_VALVE_FAULT.XV02_FAIL_TO_OPEN, FAIL_TO_CLOSE => "Valves Data".R5_VALVE_FAULT.XV02_FAIL_TO_CLOSE, status => "Valves Data".R5_XV02.STATUS)
   END_RUNG
   RUNG wire#powerrail
      Contact( "R5_DATA".R5.CTS_CMD_2 )
   END_RUNG wire#w1
   RUNG wire#powerrail
      Contact( "R5_DATA".R5.CTS_CMD_1 )
   END_RUNG wire#w1
   RUNG wire#powerrail
      Contact( "R5_DATA".R5.CTS_CMD )
   END_RUNG wire#w1
   RUNG wire#powerrail
      Contact( "R5_DATA".R5.CSV_CMD_3 )
   END_RUNG wire#w1
   RUNG wire#powerrail
      Contact( "Valves Data".R5_XV02.MCMD )
      I_Contact( "dummy".R5.Intl_2 )
   END_RUNG wire#w2
   RUNG wire#powerrail
      Contact( "Valves Data".R5_XV02.RESET )
   END_RUNG wire#w3
   RUNG wire#powerrail
      Contact( "R5_DATA".R5.Reset )
   END_RUNG wire#w3
   RUNG wire#powerrail
      I_Contact( "DI_INPUTS".R5_INPUTS_RUA.EMG_PB )
   END_RUNG wire#w4
   RUNG wire#powerrail
      Contact( "AlwaysTRUE" )
      wire#w5
      { S7_Templates := "SrcType := Int" } EQ_Contact(in1 := "Valves Data".R5_XV01.STATUS, in2 := 1)
      wire#w6
      Coil( "dummy".R5.Intl_2 )
   END_RUNG
   RUNG wire#w5
      { S7_Templates := "SrcType := Int" } EQ_Contact(in1 := "Valves Data".R5_XV03.STATUS, in2 := 1)
   END_RUNG wire#w6
   RUNG wire#w5
      { S7_Templates := "SrcType := Int" } EQ_Contact(in1 := "Valves Data".R1_XV05.STATUS, in2 := 1)
   END_RUNG wire#w6
   // the same network as SCL:
   IF "AlwaysTRUE" THEN
       #valve_R5_XV3("auto/manual" := "Valves Data"."A/M".R5,   // "valve"
                     open_auto := "R5_DATA".R5.CTS_CMD_2 OR "R5_DATA".R5.CTS_CMD_1 OR "R5_DATA".R5.CTS_CMD OR "R5_DATA".R5.CSV_CMD_3,
                     open_man := "Valves Data".R5_XV02.MCMD AND NOT "dummy".R5.Intl_2,
                     fbk_open := "A/GLR_005_XV502_OFB",
                     fbk_close := "A/GLR_005_XV502_CFB",
                     reset := "Valves Data".R5_XV02.RESET OR "R5_DATA".R5.Reset,
                     intl := NOT "DI_INPUTS".R5_INPUTS_RUA.EMG_PB,
                     Mon_En := 1,
                     mon_sp := "Valves Data".R5_XV02.MON_TIME,
                     SEMI := "Valves Data".SEMI_AUTO.R5,
                     "open/close" => "A/GLR_005_XV502_CMD",
                     FAIL_TO_OPEN => "Valves Data".R5_VALVE_FAULT.XV02_FAIL_TO_OPEN,
                     FAIL_TO_CLOSE => "Valves Data".R5_VALVE_FAULT.XV02_FAIL_TO_CLOSE,
                     status => "Valves Data".R5_XV02.STATUS);
   END_IF;
   "dummy".R5.Intl_2 := "AlwaysTRUE" AND (("Valves Data".R5_XV01.STATUS = 1) OR ("Valves Data".R5_XV03.STATUS = 1) OR ("Valves Data".R1_XV05.STATUS = 1));
END_REGION

REGION Network 47: R5_XV03
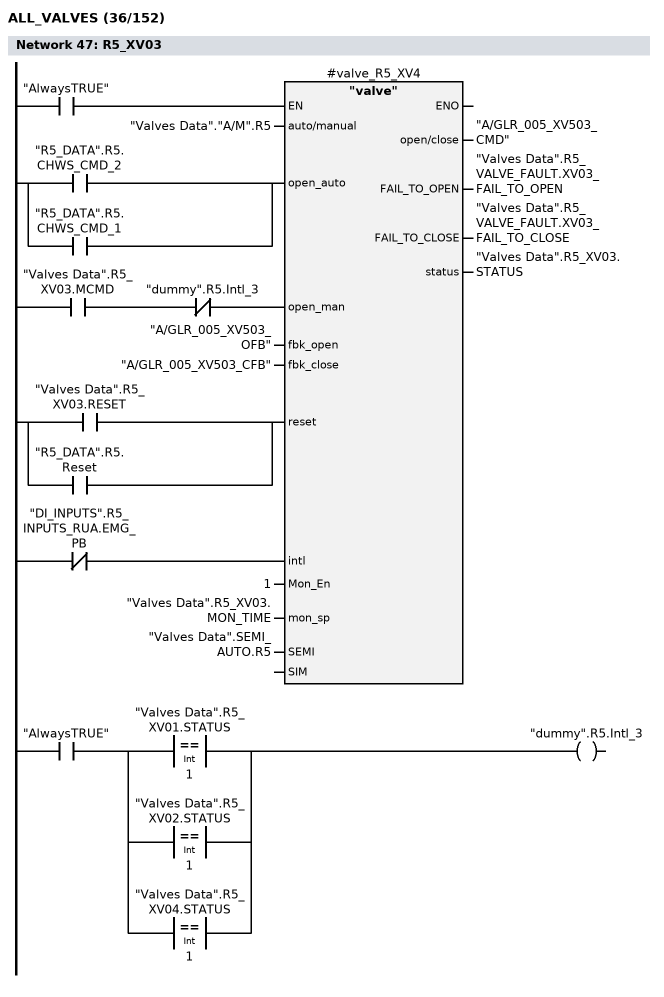
   RUNG wire#powerrail
      Contact( "AlwaysTRUE" )
      #valve_R5_XV4(open_auto := wire#w1, open_man := wire#w2, reset := wire#w3, intl := wire#w4, "auto/manual" := "Valves Data"."A/M".R5, fbk_open := "A/GLR_005_XV503_OFB", fbk_close := "A/GLR_005_XV503_CFB", Mon_En := 1, mon_sp := "Valves Data".R5_XV03.MON_TIME, SEMI := "Valves Data".SEMI_AUTO.R5, SIM :=, "open/close" => "A/GLR_005_XV503_CMD", FAIL_TO_OPEN => "Valves Data".R5_VALVE_FAULT.XV03_FAIL_TO_OPEN, FAIL_TO_CLOSE => "Valves Data".R5_VALVE_FAULT.XV03_FAIL_TO_CLOSE, status => "Valves Data".R5_XV03.STATUS)
   END_RUNG
   RUNG wire#powerrail
      Contact( "R5_DATA".R5.CHWS_CMD_2 )
   END_RUNG wire#w1
   RUNG wire#powerrail
      Contact( "R5_DATA".R5.CHWS_CMD_1 )
   END_RUNG wire#w1
   RUNG wire#powerrail
      Contact( "Valves Data".R5_XV03.MCMD )
      I_Contact( "dummy".R5.Intl_3 )
   END_RUNG wire#w2
   RUNG wire#powerrail
      Contact( "Valves Data".R5_XV03.RESET )
   END_RUNG wire#w3
   RUNG wire#powerrail
      Contact( "R5_DATA".R5.Reset )
   END_RUNG wire#w3
   RUNG wire#powerrail
      I_Contact( "DI_INPUTS".R5_INPUTS_RUA.EMG_PB )
   END_RUNG wire#w4
   RUNG wire#powerrail
      Contact( "AlwaysTRUE" )
      wire#w5
      { S7_Templates := "SrcType := Int" } EQ_Contact(in1 := "Valves Data".R5_XV01.STATUS, in2 := 1)
      wire#w6
      Coil( "dummy".R5.Intl_3 )
   END_RUNG
   RUNG wire#w5
      { S7_Templates := "SrcType := Int" } EQ_Contact(in1 := "Valves Data".R5_XV02.STATUS, in2 := 1)
   END_RUNG wire#w6
   RUNG wire#w5
      { S7_Templates := "SrcType := Int" } EQ_Contact(in1 := "Valves Data".R5_XV04.STATUS, in2 := 1)
   END_RUNG wire#w6
   // the same network as SCL:
   IF "AlwaysTRUE" THEN
       #valve_R5_XV4("auto/manual" := "Valves Data"."A/M".R5,   // "valve"
                     open_auto := "R5_DATA".R5.CHWS_CMD_2 OR "R5_DATA".R5.CHWS_CMD_1,
                     open_man := "Valves Data".R5_XV03.MCMD AND NOT "dummy".R5.Intl_3,
                     fbk_open := "A/GLR_005_XV503_OFB",
                     fbk_close := "A/GLR_005_XV503_CFB",
                     reset := "Valves Data".R5_XV03.RESET OR "R5_DATA".R5.Reset,
                     intl := NOT "DI_INPUTS".R5_INPUTS_RUA.EMG_PB,
                     Mon_En := 1,
                     mon_sp := "Valves Data".R5_XV03.MON_TIME,
                     SEMI := "Valves Data".SEMI_AUTO.R5,
                     "open/close" => "A/GLR_005_XV503_CMD",
                     FAIL_TO_OPEN => "Valves Data".R5_VALVE_FAULT.XV03_FAIL_TO_OPEN,
                     FAIL_TO_CLOSE => "Valves Data".R5_VALVE_FAULT.XV03_FAIL_TO_CLOSE,
                     status => "Valves Data".R5_XV03.STATUS);
   END_IF;
   "dummy".R5.Intl_3 := "AlwaysTRUE" AND (("Valves Data".R5_XV01.STATUS = 1) OR ("Valves Data".R5_XV02.STATUS = 1) OR ("Valves Data".R5_XV04.STATUS = 1));
END_REGION

REGION Network 48: R5_XV04
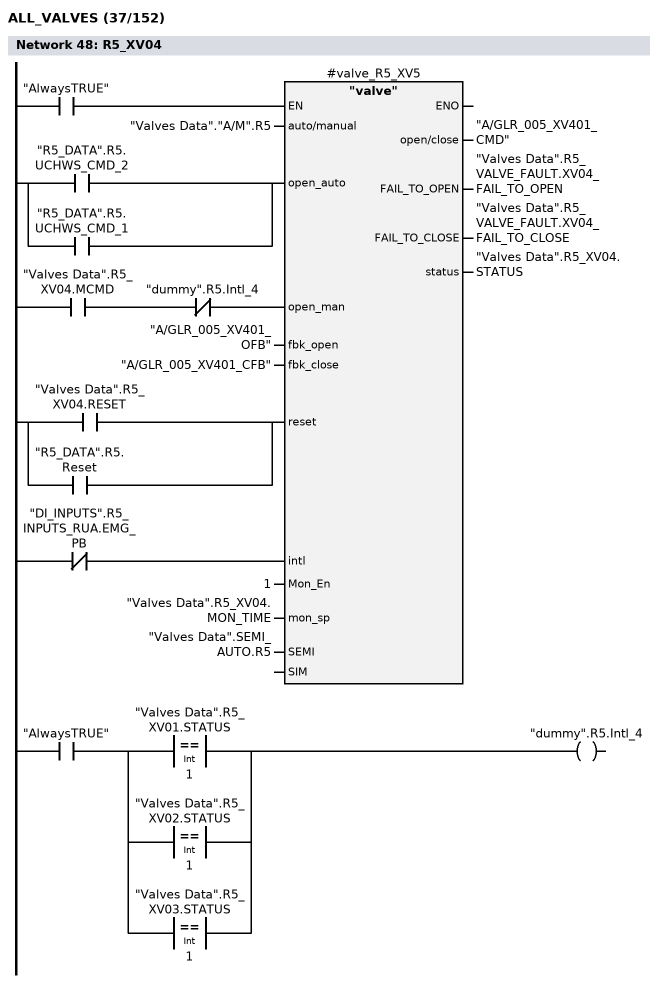
   RUNG wire#powerrail
      Contact( "AlwaysTRUE" )
      #valve_R5_XV5(open_auto := wire#w1, open_man := wire#w2, reset := wire#w3, intl := wire#w4, "auto/manual" := "Valves Data"."A/M".R5, fbk_open := "A/GLR_005_XV401_OFB", fbk_close := "A/GLR_005_XV401_CFB", Mon_En := 1, mon_sp := "Valves Data".R5_XV04.MON_TIME, SEMI := "Valves Data".SEMI_AUTO.R5, SIM :=, "open/close" => "A/GLR_005_XV401_CMD", FAIL_TO_OPEN => "Valves Data".R5_VALVE_FAULT.XV04_FAIL_TO_OPEN, FAIL_TO_CLOSE => "Valves Data".R5_VALVE_FAULT.XV04_FAIL_TO_CLOSE, status => "Valves Data".R5_XV04.STATUS)
   END_RUNG
   RUNG wire#powerrail
      Contact( "R5_DATA".R5.UCHWS_CMD_2 )
   END_RUNG wire#w1
   RUNG wire#powerrail
      Contact( "R5_DATA".R5.UCHWS_CMD_1 )
   END_RUNG wire#w1
   RUNG wire#powerrail
      Contact( "Valves Data".R5_XV04.MCMD )
      I_Contact( "dummy".R5.Intl_4 )
   END_RUNG wire#w2
   RUNG wire#powerrail
      Contact( "Valves Data".R5_XV04.RESET )
   END_RUNG wire#w3
   RUNG wire#powerrail
      Contact( "R5_DATA".R5.Reset )
   END_RUNG wire#w3
   RUNG wire#powerrail
      I_Contact( "DI_INPUTS".R5_INPUTS_RUA.EMG_PB )
   END_RUNG wire#w4
   RUNG wire#powerrail
      Contact( "AlwaysTRUE" )
      wire#w5
      { S7_Templates := "SrcType := Int" } EQ_Contact(in1 := "Valves Data".R5_XV01.STATUS, in2 := 1)
      wire#w6
      Coil( "dummy".R5.Intl_4 )
   END_RUNG
   RUNG wire#w5
      { S7_Templates := "SrcType := Int" } EQ_Contact(in1 := "Valves Data".R5_XV02.STATUS, in2 := 1)
   END_RUNG wire#w6
   RUNG wire#w5
      { S7_Templates := "SrcType := Int" } EQ_Contact(in1 := "Valves Data".R5_XV03.STATUS, in2 := 1)
   END_RUNG wire#w6
   // the same network as SCL:
   IF "AlwaysTRUE" THEN
       #valve_R5_XV5("auto/manual" := "Valves Data"."A/M".R5,   // "valve"
                     open_auto := "R5_DATA".R5.UCHWS_CMD_2 OR "R5_DATA".R5.UCHWS_CMD_1,
                     open_man := "Valves Data".R5_XV04.MCMD AND NOT "dummy".R5.Intl_4,
                     fbk_open := "A/GLR_005_XV401_OFB",
                     fbk_close := "A/GLR_005_XV401_CFB",
                     reset := "Valves Data".R5_XV04.RESET OR "R5_DATA".R5.Reset,
                     intl := NOT "DI_INPUTS".R5_INPUTS_RUA.EMG_PB,
                     Mon_En := 1,
                     mon_sp := "Valves Data".R5_XV04.MON_TIME,
                     SEMI := "Valves Data".SEMI_AUTO.R5,
                     "open/close" => "A/GLR_005_XV401_CMD",
                     FAIL_TO_OPEN => "Valves Data".R5_VALVE_FAULT.XV04_FAIL_TO_OPEN,
                     FAIL_TO_CLOSE => "Valves Data".R5_VALVE_FAULT.XV04_FAIL_TO_CLOSE,
                     status => "Valves Data".R5_XV04.STATUS);
   END_IF;
   "dummy".R5.Intl_4 := "AlwaysTRUE" AND (("Valves Data".R5_XV01.STATUS = 1) OR ("Valves Data".R5_XV02.STATUS = 1) OR ("Valves Data".R5_XV03.STATUS = 1));
END_REGION

REGION Network 49: R5_XV05
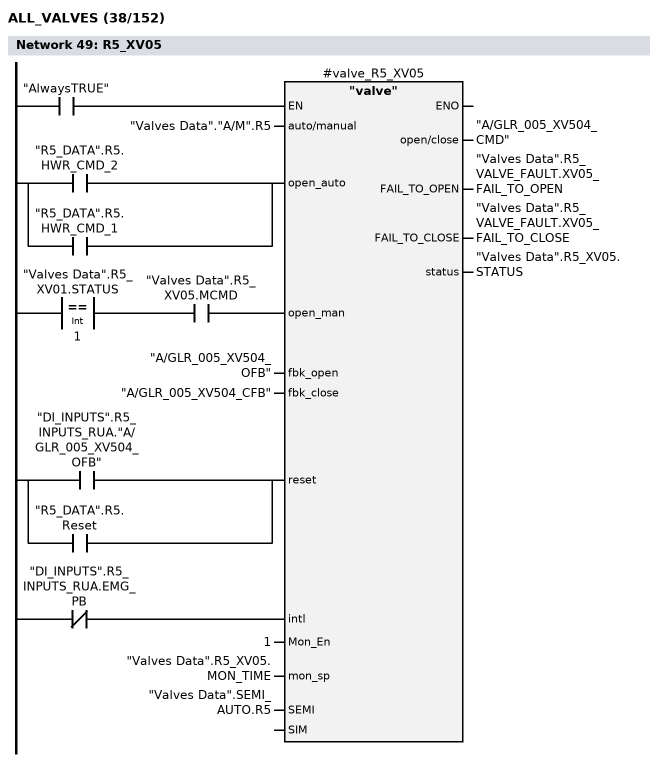
   RUNG wire#powerrail
      Contact( "AlwaysTRUE" )
      #valve_R5_XV05(open_auto := wire#w1, open_man := wire#w2, reset := wire#w3, intl := wire#w4, "auto/manual" := "Valves Data"."A/M".R5, fbk_open := "A/GLR_005_XV504_OFB", fbk_close := "A/GLR_005_XV504_CFB", Mon_En := 1, mon_sp := "Valves Data".R5_XV05.MON_TIME, SEMI := "Valves Data".SEMI_AUTO.R5, SIM :=, "open/close" => "A/GLR_005_XV504_CMD", FAIL_TO_OPEN => "Valves Data".R5_VALVE_FAULT.XV05_FAIL_TO_OPEN, FAIL_TO_CLOSE => "Valves Data".R5_VALVE_FAULT.XV05_FAIL_TO_CLOSE, status => "Valves Data".R5_XV05.STATUS)
   END_RUNG
   RUNG wire#powerrail
      Contact( "R5_DATA".R5.HWR_CMD_2 )
   END_RUNG wire#w1
   RUNG wire#powerrail
      Contact( "R5_DATA".R5.HWR_CMD_1 )
   END_RUNG wire#w1
   RUNG wire#powerrail
      { S7_Templates := "SrcType := Int" } EQ_Contact(in1 := "Valves Data".R5_XV01.STATUS, in2 := 1)
      Contact( "Valves Data".R5_XV05.MCMD )
   END_RUNG wire#w2
   RUNG wire#powerrail
      Contact( "DI_INPUTS".R5_INPUTS_RUA."A/GLR_005_XV504_OFB" )
   END_RUNG wire#w3
   RUNG wire#powerrail
      Contact( "R5_DATA".R5.Reset )
   END_RUNG wire#w3
   RUNG wire#powerrail
      I_Contact( "DI_INPUTS".R5_INPUTS_RUA.EMG_PB )
   END_RUNG wire#w4
   // the same network as SCL:
   IF "AlwaysTRUE" THEN
       #valve_R5_XV05("auto/manual" := "Valves Data"."A/M".R5,   // "valve"
                      open_auto := "R5_DATA".R5.HWR_CMD_2 OR "R5_DATA".R5.HWR_CMD_1,
                      open_man := ("Valves Data".R5_XV01.STATUS = 1) AND "Valves Data".R5_XV05.MCMD,
                      fbk_open := "A/GLR_005_XV504_OFB",
                      fbk_close := "A/GLR_005_XV504_CFB",
                      reset := "DI_INPUTS".R5_INPUTS_RUA."A/GLR_005_XV504_OFB" OR "R5_DATA".R5.Reset,
                      intl := NOT "DI_INPUTS".R5_INPUTS_RUA.EMG_PB,
                      Mon_En := 1,
                      mon_sp := "Valves Data".R5_XV05.MON_TIME,
                      SEMI := "Valves Data".SEMI_AUTO.R5,
                      "open/close" => "A/GLR_005_XV504_CMD",
                      FAIL_TO_OPEN => "Valves Data".R5_VALVE_FAULT.XV05_FAIL_TO_OPEN,
                      FAIL_TO_CLOSE => "Valves Data".R5_VALVE_FAULT.XV05_FAIL_TO_CLOSE,
                      status => "Valves Data".R5_XV05.STATUS);
   END_IF;
END_REGION

REGION Network 50: R5_XV06
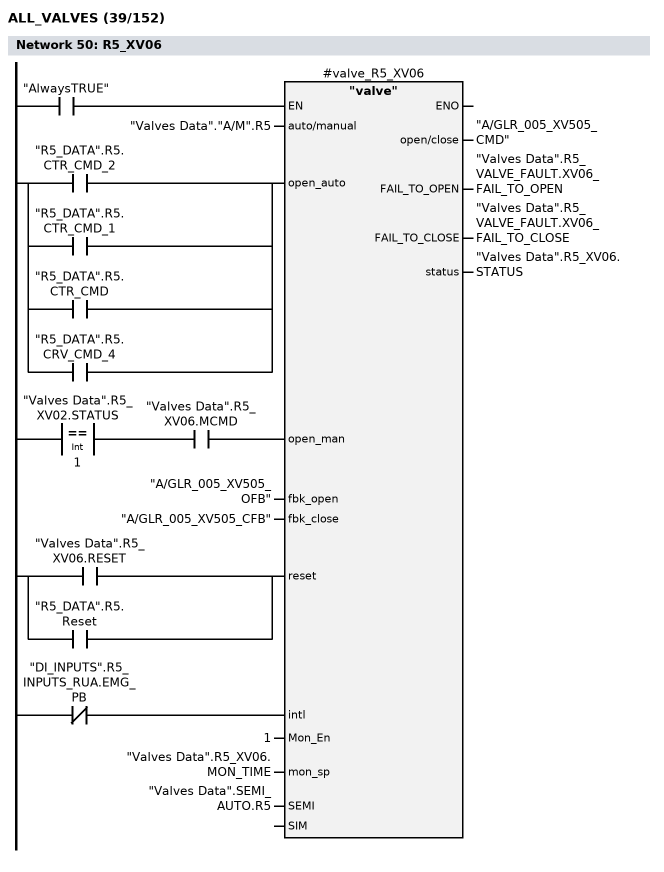
   RUNG wire#powerrail
      Contact( "AlwaysTRUE" )
      #valve_R5_XV06(open_auto := wire#w1, open_man := wire#w2, reset := wire#w3, intl := wire#w4, "auto/manual" := "Valves Data"."A/M".R5, fbk_open := "A/GLR_005_XV505_OFB", fbk_close := "A/GLR_005_XV505_CFB", Mon_En := 1, mon_sp := "Valves Data".R5_XV06.MON_TIME, SEMI := "Valves Data".SEMI_AUTO.R5, SIM :=, "open/close" => "A/GLR_005_XV505_CMD", FAIL_TO_OPEN => "Valves Data".R5_VALVE_FAULT.XV06_FAIL_TO_OPEN, FAIL_TO_CLOSE => "Valves Data".R5_VALVE_FAULT.XV06_FAIL_TO_CLOSE, status => "Valves Data".R5_XV06.STATUS)
   END_RUNG
   RUNG wire#powerrail
      Contact( "R5_DATA".R5.CTR_CMD_2 )
   END_RUNG wire#w1
   RUNG wire#powerrail
      Contact( "R5_DATA".R5.CTR_CMD_1 )
   END_RUNG wire#w1
   RUNG wire#powerrail
      Contact( "R5_DATA".R5.CTR_CMD )
   END_RUNG wire#w1
   RUNG wire#powerrail
      Contact( "R5_DATA".R5.CRV_CMD_4 )
   END_RUNG wire#w1
   RUNG wire#powerrail
      { S7_Templates := "SrcType := Int" } EQ_Contact(in1 := "Valves Data".R5_XV02.STATUS, in2 := 1)
      Contact( "Valves Data".R5_XV06.MCMD )
   END_RUNG wire#w2
   RUNG wire#powerrail
      Contact( "Valves Data".R5_XV06.RESET )
   END_RUNG wire#w3
   RUNG wire#powerrail
      Contact( "R5_DATA".R5.Reset )
   END_RUNG wire#w3
   RUNG wire#powerrail
      I_Contact( "DI_INPUTS".R5_INPUTS_RUA.EMG_PB )
   END_RUNG wire#w4
   // the same network as SCL:
   IF "AlwaysTRUE" THEN
       #valve_R5_XV06("auto/manual" := "Valves Data"."A/M".R5,   // "valve"
                      open_auto := "R5_DATA".R5.CTR_CMD_2 OR "R5_DATA".R5.CTR_CMD_1 OR "R5_DATA".R5.CTR_CMD OR "R5_DATA".R5.CRV_CMD_4,
                      open_man := ("Valves Data".R5_XV02.STATUS = 1) AND "Valves Data".R5_XV06.MCMD,
                      fbk_open := "A/GLR_005_XV505_OFB",
                      fbk_close := "A/GLR_005_XV505_CFB",
                      reset := "Valves Data".R5_XV06.RESET OR "R5_DATA".R5.Reset,
                      intl := NOT "DI_INPUTS".R5_INPUTS_RUA.EMG_PB,
                      Mon_En := 1,
                      mon_sp := "Valves Data".R5_XV06.MON_TIME,
                      SEMI := "Valves Data".SEMI_AUTO.R5,
                      "open/close" => "A/GLR_005_XV505_CMD",
                      FAIL_TO_OPEN => "Valves Data".R5_VALVE_FAULT.XV06_FAIL_TO_OPEN,
                      FAIL_TO_CLOSE => "Valves Data".R5_VALVE_FAULT.XV06_FAIL_TO_CLOSE,
                      status => "Valves Data".R5_XV06.STATUS);
   END_IF;
END_REGION

REGION Network 51: R5_XV07
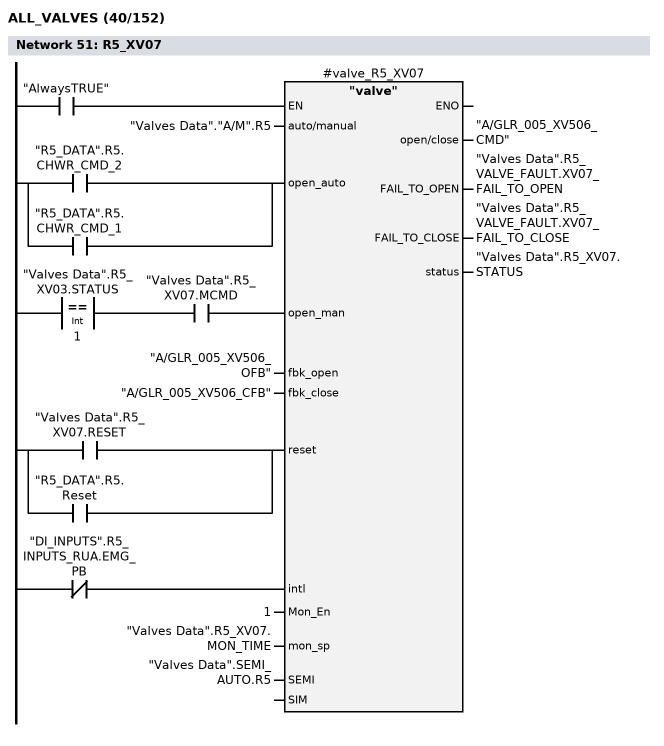
   RUNG wire#powerrail
      Contact( "AlwaysTRUE" )
      #valve_R5_XV07(open_auto := wire#w1, open_man := wire#w2, reset := wire#w3, intl := wire#w4, "auto/manual" := "Valves Data"."A/M".R5, fbk_open := "A/GLR_005_XV506_OFB", fbk_close := "A/GLR_005_XV506_CFB", Mon_En := 1, mon_sp := "Valves Data".R5_XV07.MON_TIME, SEMI := "Valves Data".SEMI_AUTO.R5, SIM :=, "open/close" => "A/GLR_005_XV506_CMD", FAIL_TO_OPEN => "Valves Data".R5_VALVE_FAULT.XV07_FAIL_TO_OPEN, FAIL_TO_CLOSE => "Valves Data".R5_VALVE_FAULT.XV07_FAIL_TO_CLOSE, status => "Valves Data".R5_XV07.STATUS)
   END_RUNG
   RUNG wire#powerrail
      Contact( "R5_DATA".R5.CHWR_CMD_2 )
   END_RUNG wire#w1
   RUNG wire#powerrail
      Contact( "R5_DATA".R5.CHWR_CMD_1 )
   END_RUNG wire#w1
   RUNG wire#powerrail
      { S7_Templates := "SrcType := Int" } EQ_Contact(in1 := "Valves Data".R5_XV03.STATUS, in2 := 1)
      Contact( "Valves Data".R5_XV07.MCMD )
   END_RUNG wire#w2
   RUNG wire#powerrail
      Contact( "Valves Data".R5_XV07.RESET )
   END_RUNG wire#w3
   RUNG wire#powerrail
      Contact( "R5_DATA".R5.Reset )
   END_RUNG wire#w3
   RUNG wire#powerrail
      I_Contact( "DI_INPUTS".R5_INPUTS_RUA.EMG_PB )
   END_RUNG wire#w4
   // the same network as SCL:
   IF "AlwaysTRUE" THEN
       #valve_R5_XV07("auto/manual" := "Valves Data"."A/M".R5,   // "valve"
                      open_auto := "R5_DATA".R5.CHWR_CMD_2 OR "R5_DATA".R5.CHWR_CMD_1,
                      open_man := ("Valves Data".R5_XV03.STATUS = 1) AND "Valves Data".R5_XV07.MCMD,
                      fbk_open := "A/GLR_005_XV506_OFB",
                      fbk_close := "A/GLR_005_XV506_CFB",
                      reset := "Valves Data".R5_XV07.RESET OR "R5_DATA".R5.Reset,
                      intl := NOT "DI_INPUTS".R5_INPUTS_RUA.EMG_PB,
                      Mon_En := 1,
                      mon_sp := "Valves Data".R5_XV07.MON_TIME,
                      SEMI := "Valves Data".SEMI_AUTO.R5,
                      "open/close" => "A/GLR_005_XV506_CMD",
                      FAIL_TO_OPEN => "Valves Data".R5_VALVE_FAULT.XV07_FAIL_TO_OPEN,
                      FAIL_TO_CLOSE => "Valves Data".R5_VALVE_FAULT.XV07_FAIL_TO_CLOSE,
                      status => "Valves Data".R5_XV07.STATUS);
   END_IF;
END_REGION

REGION Network 52: R5_XV08
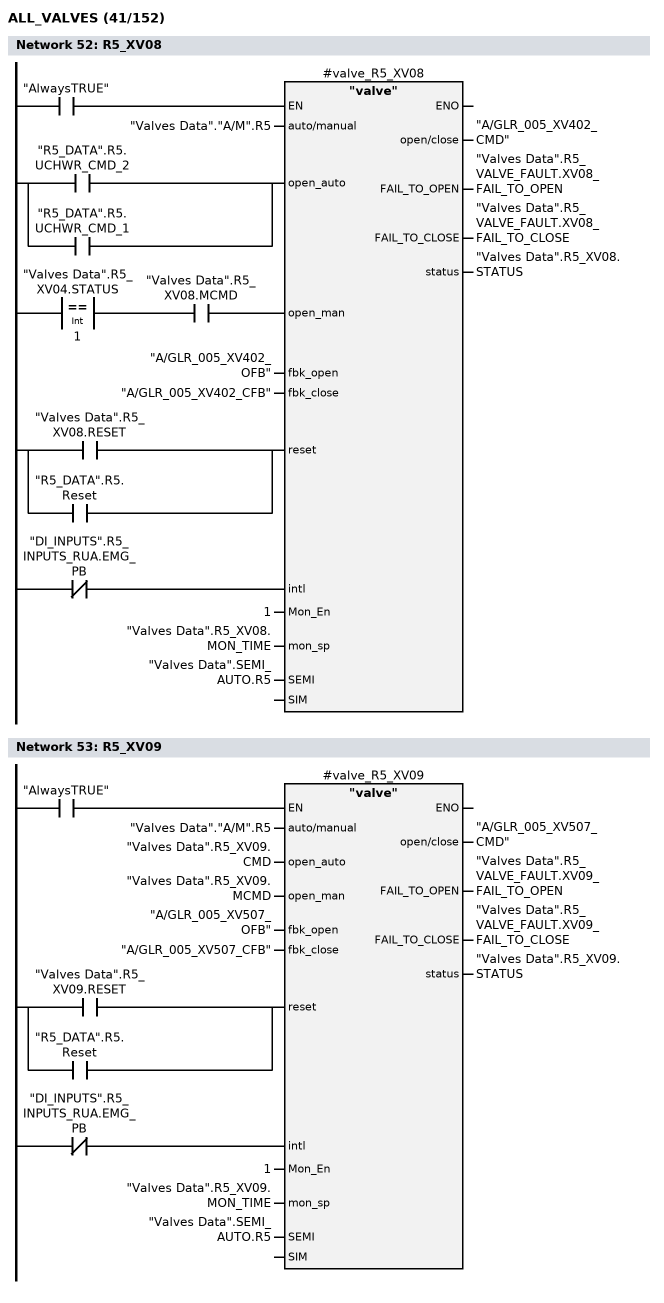
   RUNG wire#powerrail
      Contact( "AlwaysTRUE" )
      #valve_R5_XV08(open_auto := wire#w1, open_man := wire#w2, reset := wire#w3, intl := wire#w4, "auto/manual" := "Valves Data"."A/M".R5, fbk_open := "A/GLR_005_XV402_OFB", fbk_close := "A/GLR_005_XV402_CFB", Mon_En := 1, mon_sp := "Valves Data".R5_XV08.MON_TIME, SEMI := "Valves Data".SEMI_AUTO.R5, SIM :=, "open/close" => "A/GLR_005_XV402_CMD", FAIL_TO_OPEN => "Valves Data".R5_VALVE_FAULT.XV08_FAIL_TO_OPEN, FAIL_TO_CLOSE => "Valves Data".R5_VALVE_FAULT.XV08_FAIL_TO_CLOSE, status => "Valves Data".R5_XV08.STATUS)
   END_RUNG
   RUNG wire#powerrail
      Contact( "R5_DATA".R5.UCHWR_CMD_2 )
   END_RUNG wire#w1
   RUNG wire#powerrail
      Contact( "R5_DATA".R5.UCHWR_CMD_1 )
   END_RUNG wire#w1
   RUNG wire#powerrail
      { S7_Templates := "SrcType := Int" } EQ_Contact(in1 := "Valves Data".R5_XV04.STATUS, in2 := 1)
      Contact( "Valves Data".R5_XV08.MCMD )
   END_RUNG wire#w2
   RUNG wire#powerrail
      Contact( "Valves Data".R5_XV08.RESET )
   END_RUNG wire#w3
   RUNG wire#powerrail
      Contact( "R5_DATA".R5.Reset )
   END_RUNG wire#w3
   RUNG wire#powerrail
      I_Contact( "DI_INPUTS".R5_INPUTS_RUA.EMG_PB )
   END_RUNG wire#w4
   // the same network as SCL:
   IF "AlwaysTRUE" THEN
       #valve_R5_XV08("auto/manual" := "Valves Data"."A/M".R5,   // "valve"
                      open_auto := "R5_DATA".R5.UCHWR_CMD_2 OR "R5_DATA".R5.UCHWR_CMD_1,
                      open_man := ("Valves Data".R5_XV04.STATUS = 1) AND "Valves Data".R5_XV08.MCMD,
                      fbk_open := "A/GLR_005_XV402_OFB",
                      fbk_close := "A/GLR_005_XV402_CFB",
                      reset := "Valves Data".R5_XV08.RESET OR "R5_DATA".R5.Reset,
                      intl := NOT "DI_INPUTS".R5_INPUTS_RUA.EMG_PB,
                      Mon_En := 1,
                      mon_sp := "Valves Data".R5_XV08.MON_TIME,
                      SEMI := "Valves Data".SEMI_AUTO.R5,
                      "open/close" => "A/GLR_005_XV402_CMD",
                      FAIL_TO_OPEN => "Valves Data".R5_VALVE_FAULT.XV08_FAIL_TO_OPEN,
                      FAIL_TO_CLOSE => "Valves Data".R5_VALVE_FAULT.XV08_FAIL_TO_CLOSE,
                      status => "Valves Data".R5_XV08.STATUS);
   END_IF;
END_REGION

REGION Network 53: R5_XV09
   RUNG wire#powerrail
      Contact( "AlwaysTRUE" )
      #valve_R5_XV09(reset := wire#w1, intl := wire#w2, "auto/manual" := "Valves Data"."A/M".R5, open_auto := "Valves Data".R5_XV09.CMD, open_man := "Valves Data".R5_XV09.MCMD, fbk_open := "A/GLR_005_XV507_OFB", fbk_close := "A/GLR_005_XV507_CFB", Mon_En := 1, mon_sp := "Valves Data".R5_XV09.MON_TIME, SEMI := "Valves Data".SEMI_AUTO.R5, SIM :=, "open/close" => "A/GLR_005_XV507_CMD", FAIL_TO_OPEN => "Valves Data".R5_VALVE_FAULT.XV09_FAIL_TO_OPEN, FAIL_TO_CLOSE => "Valves Data".R5_VALVE_FAULT.XV09_FAIL_TO_CLOSE, status => "Valves Data".R5_XV09.STATUS)
   END_RUNG
   RUNG wire#powerrail
      Contact( "Valves Data".R5_XV09.RESET )
   END_RUNG wire#w1
   RUNG wire#powerrail
      Contact( "R5_DATA".R5.Reset )
   END_RUNG wire#w1
   RUNG wire#powerrail
      I_Contact( "DI_INPUTS".R5_INPUTS_RUA.EMG_PB )
   END_RUNG wire#w2
   // the same network as SCL:
   IF "AlwaysTRUE" THEN
       #valve_R5_XV09("auto/manual" := "Valves Data"."A/M".R5,   // "valve"
                      open_auto := "Valves Data".R5_XV09.CMD,
                      open_man := "Valves Data".R5_XV09.MCMD,
                      fbk_open := "A/GLR_005_XV507_OFB",
                      fbk_close := "A/GLR_005_XV507_CFB",
                      reset := "Valves Data".R5_XV09.RESET OR "R5_DATA".R5.Reset,
                      intl := NOT "DI_INPUTS".R5_INPUTS_RUA.EMG_PB,
                      Mon_En := 1,
                      mon_sp := "Valves Data".R5_XV09.MON_TIME,
                      SEMI := "Valves Data".SEMI_AUTO.R5,
                      "open/close" => "A/GLR_005_XV507_CMD",
                      FAIL_TO_OPEN => "Valves Data".R5_VALVE_FAULT.XV09_FAIL_TO_OPEN,
                      FAIL_TO_CLOSE => "Valves Data".R5_VALVE_FAULT.XV09_FAIL_TO_CLOSE,
                      status => "Valves Data".R5_XV09.STATUS);
   END_IF;
END_REGION

REGION Network 54: R5_XV10
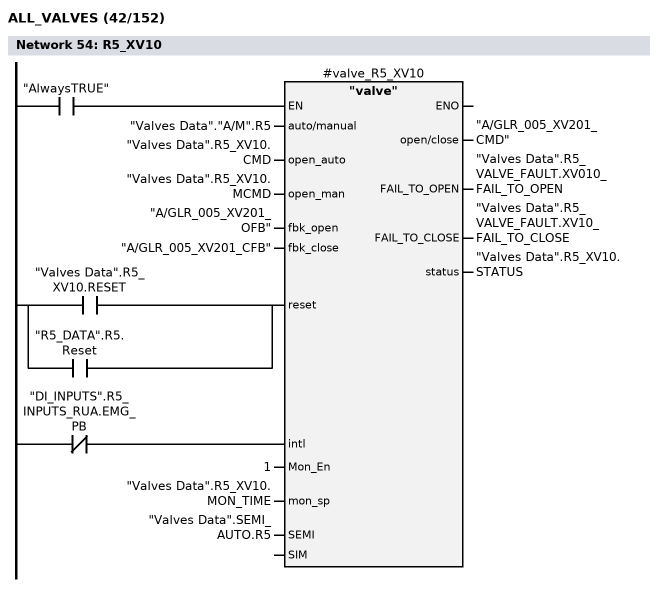
   RUNG wire#powerrail
      Contact( "AlwaysTRUE" )
      #valve_R5_XV10(reset := wire#w1, intl := wire#w2, "auto/manual" := "Valves Data"."A/M".R5, open_auto := "Valves Data".R5_XV10.CMD, open_man := "Valves Data".R5_XV10.MCMD, fbk_open := "A/GLR_005_XV201_OFB", fbk_close := "A/GLR_005_XV201_CFB", Mon_En := 1, mon_sp := "Valves Data".R5_XV10.MON_TIME, SEMI := "Valves Data".SEMI_AUTO.R5, SIM :=, "open/close" => "A/GLR_005_XV201_CMD", FAIL_TO_OPEN => "Valves Data".R5_VALVE_FAULT.XV010_FAIL_TO_OPEN, FAIL_TO_CLOSE => "Valves Data".R5_VALVE_FAULT.XV10_FAIL_TO_CLOSE, status => "Valves Data".R5_XV10.STATUS)
   END_RUNG
   RUNG wire#powerrail
      Contact( "Valves Data".R5_XV10.RESET )
   END_RUNG wire#w1
   RUNG wire#powerrail
      Contact( "R5_DATA".R5.Reset )
   END_RUNG wire#w1
   RUNG wire#powerrail
      I_Contact( "DI_INPUTS".R5_INPUTS_RUA.EMG_PB )
   END_RUNG wire#w2
   // the same network as SCL:
   IF "AlwaysTRUE" THEN
       #valve_R5_XV10("auto/manual" := "Valves Data"."A/M".R5,   // "valve"
                      open_auto := "Valves Data".R5_XV10.CMD,
                      open_man := "Valves Data".R5_XV10.MCMD,
                      fbk_open := "A/GLR_005_XV201_OFB",
                      fbk_close := "A/GLR_005_XV201_CFB",
                      reset := "Valves Data".R5_XV10.RESET OR "R5_DATA".R5.Reset,
                      intl := NOT "DI_INPUTS".R5_INPUTS_RUA.EMG_PB,
                      Mon_En := 1,
                      mon_sp := "Valves Data".R5_XV10.MON_TIME,
                      SEMI := "Valves Data".SEMI_AUTO.R5,
                      "open/close" => "A/GLR_005_XV201_CMD",
                      FAIL_TO_OPEN => "Valves Data".R5_VALVE_FAULT.XV010_FAIL_TO_OPEN,
                      FAIL_TO_CLOSE => "Valves Data".R5_VALVE_FAULT.XV10_FAIL_TO_CLOSE,
                      status => "Valves Data".R5_XV10.STATUS);
   END_IF;
END_REGION

REGION Network 55: ****REACTOR_06****
END_REGION

REGION Network 56: R6_XV01
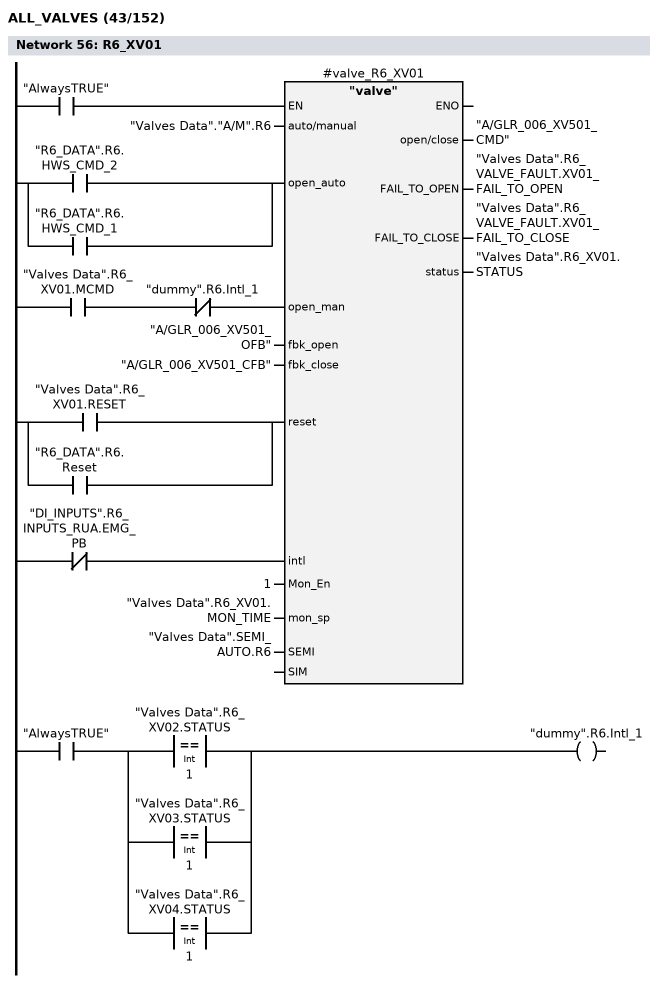
   RUNG wire#powerrail
      Contact( "AlwaysTRUE" )
      #valve_R6_XV01(open_auto := wire#w1, open_man := wire#w2, reset := wire#w3, intl := wire#w4, "auto/manual" := "Valves Data"."A/M".R6, fbk_open := "A/GLR_006_XV501_OFB", fbk_close := "A/GLR_006_XV501_CFB", Mon_En := 1, mon_sp := "Valves Data".R6_XV01.MON_TIME, SEMI := "Valves Data".SEMI_AUTO.R6, SIM :=, "open/close" => "A/GLR_006_XV501_CMD", FAIL_TO_OPEN => "Valves Data".R6_VALVE_FAULT.XV01_FAIL_TO_OPEN, FAIL_TO_CLOSE => "Valves Data".R6_VALVE_FAULT.XV01_FAIL_TO_CLOSE, status => "Valves Data".R6_XV01.STATUS)
   END_RUNG
   RUNG wire#powerrail
      Contact( "R6_DATA".R6.HWS_CMD_2 )
   END_RUNG wire#w1
   RUNG wire#powerrail
      Contact( "R6_DATA".R6.HWS_CMD_1 )
   END_RUNG wire#w1
   RUNG wire#powerrail
      Contact( "Valves Data".R6_XV01.MCMD )
      I_Contact( "dummy".R6.Intl_1 )
   END_RUNG wire#w2
   RUNG wire#powerrail
      Contact( "Valves Data".R6_XV01.RESET )
   END_RUNG wire#w3
   RUNG wire#powerrail
      Contact( "R6_DATA".R6.Reset )
   END_RUNG wire#w3
   RUNG wire#powerrail
      I_Contact( "DI_INPUTS".R6_INPUTS_RUA.EMG_PB )
   END_RUNG wire#w4
   RUNG wire#powerrail
      Contact( "AlwaysTRUE" )
      wire#w5
      { S7_Templates := "SrcType := Int" } EQ_Contact(in1 := "Valves Data".R6_XV02.STATUS, in2 := 1)
      wire#w6
      Coil( "dummy".R6.Intl_1 )
   END_RUNG
   RUNG wire#w5
      { S7_Templates := "SrcType := Int" } EQ_Contact(in1 := "Valves Data".R6_XV03.STATUS, in2 := 1)
   END_RUNG wire#w6
   RUNG wire#w5
      { S7_Templates := "SrcType := Int" } EQ_Contact(in1 := "Valves Data".R6_XV04.STATUS, in2 := 1)
   END_RUNG wire#w6
   // the same network as SCL:
   IF "AlwaysTRUE" THEN
       #valve_R6_XV01("auto/manual" := "Valves Data"."A/M".R6,   // "valve"
                      open_auto := "R6_DATA".R6.HWS_CMD_2 OR "R6_DATA".R6.HWS_CMD_1,
                      open_man := "Valves Data".R6_XV01.MCMD AND NOT "dummy".R6.Intl_1,
                      fbk_open := "A/GLR_006_XV501_OFB",
                      fbk_close := "A/GLR_006_XV501_CFB",
                      reset := "Valves Data".R6_XV01.RESET OR "R6_DATA".R6.Reset,
                      intl := NOT "DI_INPUTS".R6_INPUTS_RUA.EMG_PB,
                      Mon_En := 1,
                      mon_sp := "Valves Data".R6_XV01.MON_TIME,
                      SEMI := "Valves Data".SEMI_AUTO.R6,
                      "open/close" => "A/GLR_006_XV501_CMD",
                      FAIL_TO_OPEN => "Valves Data".R6_VALVE_FAULT.XV01_FAIL_TO_OPEN,
                      FAIL_TO_CLOSE => "Valves Data".R6_VALVE_FAULT.XV01_FAIL_TO_CLOSE,
                      status => "Valves Data".R6_XV01.STATUS);
   END_IF;
   "dummy".R6.Intl_1 := "AlwaysTRUE" AND (("Valves Data".R6_XV02.STATUS = 1) OR ("Valves Data".R6_XV03.STATUS = 1) OR ("Valves Data".R6_XV04.STATUS = 1));
END_REGION

REGION Network 57: R6_XV02
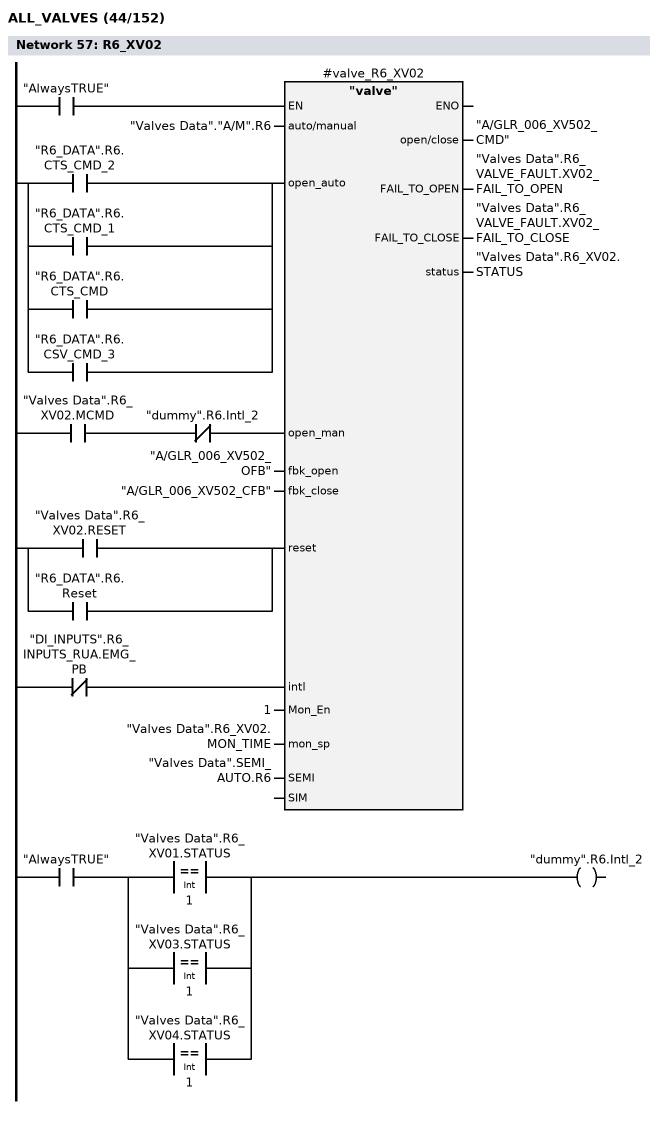
   RUNG wire#powerrail
      Contact( "AlwaysTRUE" )
      #valve_R6_XV02(open_auto := wire#w1, open_man := wire#w2, reset := wire#w3, intl := wire#w4, "auto/manual" := "Valves Data"."A/M".R6, fbk_open := "A/GLR_006_XV502_OFB", fbk_close := "A/GLR_006_XV502_CFB", Mon_En := 1, mon_sp := "Valves Data".R6_XV02.MON_TIME, SEMI := "Valves Data".SEMI_AUTO.R6, SIM :=, "open/close" => "A/GLR_006_XV502_CMD", FAIL_TO_OPEN => "Valves Data".R6_VALVE_FAULT.XV02_FAIL_TO_OPEN, FAIL_TO_CLOSE => "Valves Data".R6_VALVE_FAULT.XV02_FAIL_TO_CLOSE, status => "Valves Data".R6_XV02.STATUS)
   END_RUNG
   RUNG wire#powerrail
      Contact( "R6_DATA".R6.CTS_CMD_2 )
   END_RUNG wire#w1
   RUNG wire#powerrail
      Contact( "R6_DATA".R6.CTS_CMD_1 )
   END_RUNG wire#w1
   RUNG wire#powerrail
      Contact( "R6_DATA".R6.CTS_CMD )
   END_RUNG wire#w1
   RUNG wire#powerrail
      Contact( "R6_DATA".R6.CSV_CMD_3 )
   END_RUNG wire#w1
   RUNG wire#powerrail
      Contact( "Valves Data".R6_XV02.MCMD )
      I_Contact( "dummy".R6.Intl_2 )
   END_RUNG wire#w2
   RUNG wire#powerrail
      Contact( "Valves Data".R6_XV02.RESET )
   END_RUNG wire#w3
   RUNG wire#powerrail
      Contact( "R6_DATA".R6.Reset )
   END_RUNG wire#w3
   RUNG wire#powerrail
      I_Contact( "DI_INPUTS".R6_INPUTS_RUA.EMG_PB )
   END_RUNG wire#w4
   RUNG wire#powerrail
      Contact( "AlwaysTRUE" )
      wire#w5
      { S7_Templates := "SrcType := Int" } EQ_Contact(in1 := "Valves Data".R6_XV01.STATUS, in2 := 1)
      wire#w6
      Coil( "dummy".R6.Intl_2 )
   END_RUNG
   RUNG wire#w5
      { S7_Templates := "SrcType := Int" } EQ_Contact(in1 := "Valves Data".R6_XV03.STATUS, in2 := 1)
   END_RUNG wire#w6
   RUNG wire#w5
      { S7_Templates := "SrcType := Int" } EQ_Contact(in1 := "Valves Data".R6_XV04.STATUS, in2 := 1)
   END_RUNG wire#w6
   // the same network as SCL:
   IF "AlwaysTRUE" THEN
       #valve_R6_XV02("auto/manual" := "Valves Data"."A/M".R6,   // "valve"
                      open_auto := "R6_DATA".R6.CTS_CMD_2 OR "R6_DATA".R6.CTS_CMD_1 OR "R6_DATA".R6.CTS_CMD OR "R6_DATA".R6.CSV_CMD_3,
                      open_man := "Valves Data".R6_XV02.MCMD AND NOT "dummy".R6.Intl_2,
                      fbk_open := "A/GLR_006_XV502_OFB",
                      fbk_close := "A/GLR_006_XV502_CFB",
                      reset := "Valves Data".R6_XV02.RESET OR "R6_DATA".R6.Reset,
                      intl := NOT "DI_INPUTS".R6_INPUTS_RUA.EMG_PB,
                      Mon_En := 1,
                      mon_sp := "Valves Data".R6_XV02.MON_TIME,
                      SEMI := "Valves Data".SEMI_AUTO.R6,
                      "open/close" => "A/GLR_006_XV502_CMD",
                      FAIL_TO_OPEN => "Valves Data".R6_VALVE_FAULT.XV02_FAIL_TO_OPEN,
                      FAIL_TO_CLOSE => "Valves Data".R6_VALVE_FAULT.XV02_FAIL_TO_CLOSE,
                      status => "Valves Data".R6_XV02.STATUS);
   END_IF;
   "dummy".R6.Intl_2 := "AlwaysTRUE" AND (("Valves Data".R6_XV01.STATUS = 1) OR ("Valves Data".R6_XV03.STATUS = 1) OR ("Valves Data".R6_XV04.STATUS = 1));
END_REGION

REGION Network 58: R6_XV03
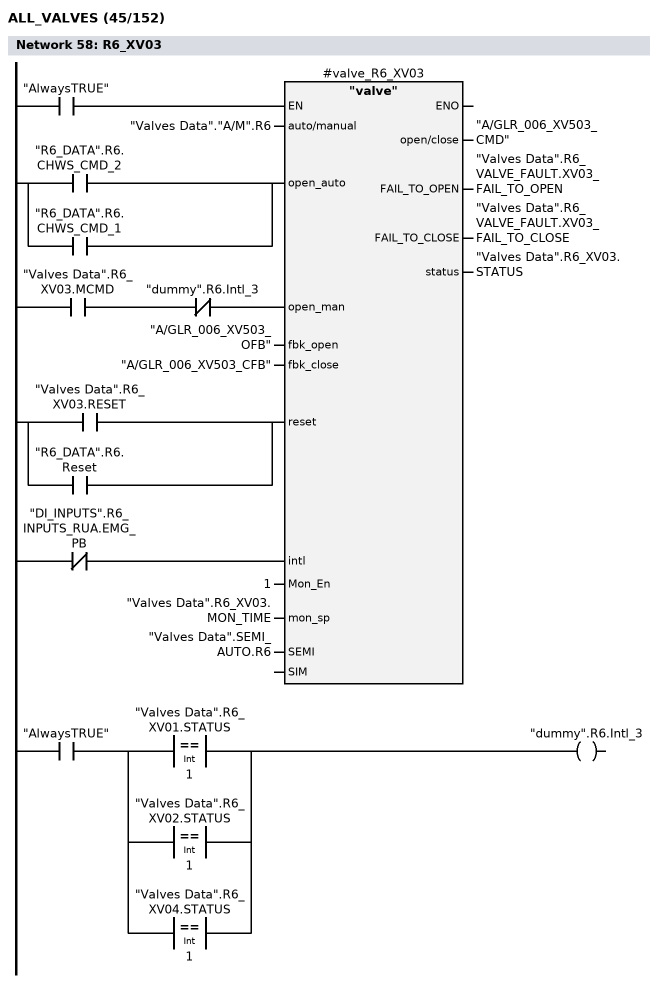
   RUNG wire#powerrail
      Contact( "AlwaysTRUE" )
      #valve_R6_XV03(open_auto := wire#w1, open_man := wire#w2, reset := wire#w3, intl := wire#w4, "auto/manual" := "Valves Data"."A/M".R6, fbk_open := "A/GLR_006_XV503_OFB", fbk_close := "A/GLR_006_XV503_CFB", Mon_En := 1, mon_sp := "Valves Data".R6_XV03.MON_TIME, SEMI := "Valves Data".SEMI_AUTO.R6, SIM :=, "open/close" => "A/GLR_006_XV503_CMD", FAIL_TO_OPEN => "Valves Data".R6_VALVE_FAULT.XV03_FAIL_TO_OPEN, FAIL_TO_CLOSE => "Valves Data".R6_VALVE_FAULT.XV03_FAIL_TO_CLOSE, status => "Valves Data".R6_XV03.STATUS)
   END_RUNG
   RUNG wire#powerrail
      Contact( "R6_DATA".R6.CHWS_CMD_2 )
   END_RUNG wire#w1
   RUNG wire#powerrail
      Contact( "R6_DATA".R6.CHWS_CMD_1 )
   END_RUNG wire#w1
   RUNG wire#powerrail
      Contact( "Valves Data".R6_XV03.MCMD )
      I_Contact( "dummy".R6.Intl_3 )
   END_RUNG wire#w2
   RUNG wire#powerrail
      Contact( "Valves Data".R6_XV03.RESET )
   END_RUNG wire#w3
   RUNG wire#powerrail
      Contact( "R6_DATA".R6.Reset )
   END_RUNG wire#w3
   RUNG wire#powerrail
      I_Contact( "DI_INPUTS".R6_INPUTS_RUA.EMG_PB )
   END_RUNG wire#w4
   RUNG wire#powerrail
      Contact( "AlwaysTRUE" )
      wire#w5
      { S7_Templates := "SrcType := Int" } EQ_Contact(in1 := "Valves Data".R6_XV01.STATUS, in2 := 1)
      wire#w6
      Coil( "dummy".R6.Intl_3 )
   END_RUNG
   RUNG wire#w5
      { S7_Templates := "SrcType := Int" } EQ_Contact(in1 := "Valves Data".R6_XV02.STATUS, in2 := 1)
   END_RUNG wire#w6
   RUNG wire#w5
      { S7_Templates := "SrcType := Int" } EQ_Contact(in1 := "Valves Data".R6_XV04.STATUS, in2 := 1)
   END_RUNG wire#w6
   // the same network as SCL:
   IF "AlwaysTRUE" THEN
       #valve_R6_XV03("auto/manual" := "Valves Data"."A/M".R6,   // "valve"
                      open_auto := "R6_DATA".R6.CHWS_CMD_2 OR "R6_DATA".R6.CHWS_CMD_1,
                      open_man := "Valves Data".R6_XV03.MCMD AND NOT "dummy".R6.Intl_3,
                      fbk_open := "A/GLR_006_XV503_OFB",
                      fbk_close := "A/GLR_006_XV503_CFB",
                      reset := "Valves Data".R6_XV03.RESET OR "R6_DATA".R6.Reset,
                      intl := NOT "DI_INPUTS".R6_INPUTS_RUA.EMG_PB,
                      Mon_En := 1,
                      mon_sp := "Valves Data".R6_XV03.MON_TIME,
                      SEMI := "Valves Data".SEMI_AUTO.R6,
                      "open/close" => "A/GLR_006_XV503_CMD",
                      FAIL_TO_OPEN => "Valves Data".R6_VALVE_FAULT.XV03_FAIL_TO_OPEN,
                      FAIL_TO_CLOSE => "Valves Data".R6_VALVE_FAULT.XV03_FAIL_TO_CLOSE,
                      status => "Valves Data".R6_XV03.STATUS);
   END_IF;
   "dummy".R6.Intl_3 := "AlwaysTRUE" AND (("Valves Data".R6_XV01.STATUS = 1) OR ("Valves Data".R6_XV02.STATUS = 1) OR ("Valves Data".R6_XV04.STATUS = 1));
END_REGION

REGION Network 59: R6_XV04
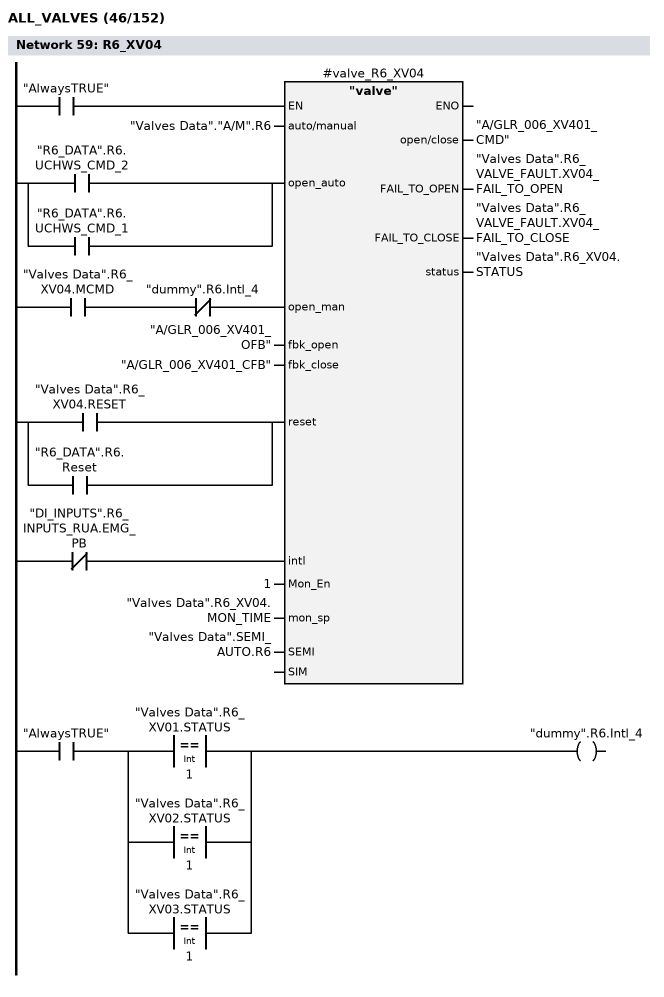
   RUNG wire#powerrail
      Contact( "AlwaysTRUE" )
      #valve_R6_XV04(open_auto := wire#w1, open_man := wire#w2, reset := wire#w3, intl := wire#w4, "auto/manual" := "Valves Data"."A/M".R6, fbk_open := "A/GLR_006_XV401_OFB", fbk_close := "A/GLR_006_XV401_CFB", Mon_En := 1, mon_sp := "Valves Data".R6_XV04.MON_TIME, SEMI := "Valves Data".SEMI_AUTO.R6, SIM :=, "open/close" => "A/GLR_006_XV401_CMD", FAIL_TO_OPEN => "Valves Data".R6_VALVE_FAULT.XV04_FAIL_TO_OPEN, FAIL_TO_CLOSE => "Valves Data".R6_VALVE_FAULT.XV04_FAIL_TO_CLOSE, status => "Valves Data".R6_XV04.STATUS)
   END_RUNG
   RUNG wire#powerrail
      Contact( "R6_DATA".R6.UCHWS_CMD_2 )
   END_RUNG wire#w1
   RUNG wire#powerrail
      Contact( "R6_DATA".R6.UCHWS_CMD_1 )
   END_RUNG wire#w1
   RUNG wire#powerrail
      Contact( "Valves Data".R6_XV04.MCMD )
      I_Contact( "dummy".R6.Intl_4 )
   END_RUNG wire#w2
   RUNG wire#powerrail
      Contact( "Valves Data".R6_XV04.RESET )
   END_RUNG wire#w3
   RUNG wire#powerrail
      Contact( "R6_DATA".R6.Reset )
   END_RUNG wire#w3
   RUNG wire#powerrail
      I_Contact( "DI_INPUTS".R6_INPUTS_RUA.EMG_PB )
   END_RUNG wire#w4
   RUNG wire#powerrail
      Contact( "AlwaysTRUE" )
      wire#w5
      { S7_Templates := "SrcType := Int" } EQ_Contact(in1 := "Valves Data".R6_XV01.STATUS, in2 := 1)
      wire#w6
      Coil( "dummy".R6.Intl_4 )
   END_RUNG
   RUNG wire#w5
      { S7_Templates := "SrcType := Int" } EQ_Contact(in1 := "Valves Data".R6_XV02.STATUS, in2 := 1)
   END_RUNG wire#w6
   RUNG wire#w5
      { S7_Templates := "SrcType := Int" } EQ_Contact(in1 := "Valves Data".R6_XV03.STATUS, in2 := 1)
   END_RUNG wire#w6
   // the same network as SCL:
   IF "AlwaysTRUE" THEN
       #valve_R6_XV04("auto/manual" := "Valves Data"."A/M".R6,   // "valve"
                      open_auto := "R6_DATA".R6.UCHWS_CMD_2 OR "R6_DATA".R6.UCHWS_CMD_1,
                      open_man := "Valves Data".R6_XV04.MCMD AND NOT "dummy".R6.Intl_4,
                      fbk_open := "A/GLR_006_XV401_OFB",
                      fbk_close := "A/GLR_006_XV401_CFB",
                      reset := "Valves Data".R6_XV04.RESET OR "R6_DATA".R6.Reset,
                      intl := NOT "DI_INPUTS".R6_INPUTS_RUA.EMG_PB,
                      Mon_En := 1,
                      mon_sp := "Valves Data".R6_XV04.MON_TIME,
                      SEMI := "Valves Data".SEMI_AUTO.R6,
                      "open/close" => "A/GLR_006_XV401_CMD",
                      FAIL_TO_OPEN => "Valves Data".R6_VALVE_FAULT.XV04_FAIL_TO_OPEN,
                      FAIL_TO_CLOSE => "Valves Data".R6_VALVE_FAULT.XV04_FAIL_TO_CLOSE,
                      status => "Valves Data".R6_XV04.STATUS);
   END_IF;
   "dummy".R6.Intl_4 := "AlwaysTRUE" AND (("Valves Data".R6_XV01.STATUS = 1) OR ("Valves Data".R6_XV02.STATUS = 1) OR ("Valves Data".R6_XV03.STATUS = 1));
END_REGION

REGION Network 60: R6_XV05
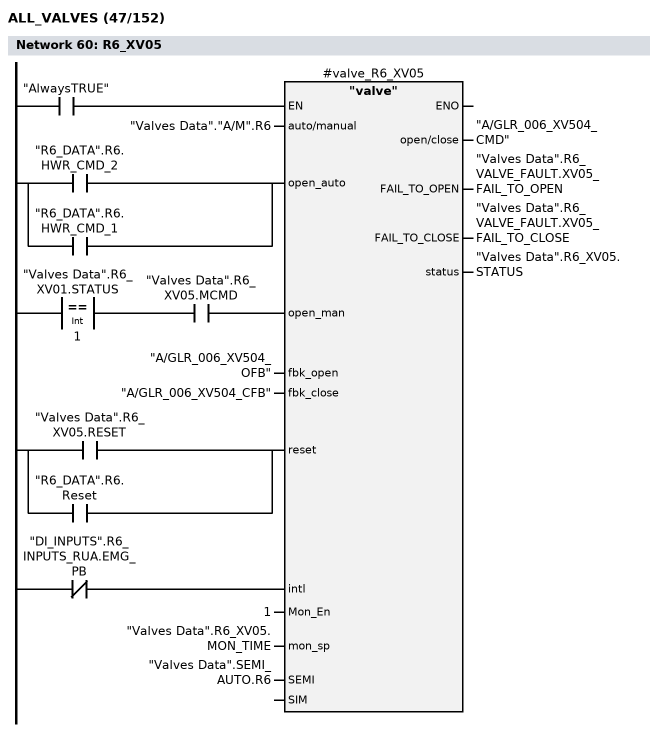
   RUNG wire#powerrail
      Contact( "AlwaysTRUE" )
      #valve_R6_XV05(open_auto := wire#w1, open_man := wire#w2, reset := wire#w3, intl := wire#w4, "auto/manual" := "Valves Data"."A/M".R6, fbk_open := "A/GLR_006_XV504_OFB", fbk_close := "A/GLR_006_XV504_CFB", Mon_En := 1, mon_sp := "Valves Data".R6_XV05.MON_TIME, SEMI := "Valves Data".SEMI_AUTO.R6, SIM :=, "open/close" => "A/GLR_006_XV504_CMD", FAIL_TO_OPEN => "Valves Data".R6_VALVE_FAULT.XV05_FAIL_TO_OPEN, FAIL_TO_CLOSE => "Valves Data".R6_VALVE_FAULT.XV05_FAIL_TO_CLOSE, status => "Valves Data".R6_XV05.STATUS)
   END_RUNG
   RUNG wire#powerrail
      Contact( "R6_DATA".R6.HWR_CMD_2 )
   END_RUNG wire#w1
   RUNG wire#powerrail
      Contact( "R6_DATA".R6.HWR_CMD_1 )
   END_RUNG wire#w1
   RUNG wire#powerrail
      { S7_Templates := "SrcType := Int" } EQ_Contact(in1 := "Valves Data".R6_XV01.STATUS, in2 := 1)
      Contact( "Valves Data".R6_XV05.MCMD )
   END_RUNG wire#w2
   RUNG wire#powerrail
      Contact( "Valves Data".R6_XV05.RESET )
   END_RUNG wire#w3
   RUNG wire#powerrail
      Contact( "R6_DATA".R6.Reset )
   END_RUNG wire#w3
   RUNG wire#powerrail
      I_Contact( "DI_INPUTS".R6_INPUTS_RUA.EMG_PB )
   END_RUNG wire#w4
   // the same network as SCL:
   IF "AlwaysTRUE" THEN
       #valve_R6_XV05("auto/manual" := "Valves Data"."A/M".R6,   // "valve"
                      open_auto := "R6_DATA".R6.HWR_CMD_2 OR "R6_DATA".R6.HWR_CMD_1,
                      open_man := ("Valves Data".R6_XV01.STATUS = 1) AND "Valves Data".R6_XV05.MCMD,
                      fbk_open := "A/GLR_006_XV504_OFB",
                      fbk_close := "A/GLR_006_XV504_CFB",
                      reset := "Valves Data".R6_XV05.RESET OR "R6_DATA".R6.Reset,
                      intl := NOT "DI_INPUTS".R6_INPUTS_RUA.EMG_PB,
                      Mon_En := 1,
                      mon_sp := "Valves Data".R6_XV05.MON_TIME,
                      SEMI := "Valves Data".SEMI_AUTO.R6,
                      "open/close" => "A/GLR_006_XV504_CMD",
                      FAIL_TO_OPEN => "Valves Data".R6_VALVE_FAULT.XV05_FAIL_TO_OPEN,
                      FAIL_TO_CLOSE => "Valves Data".R6_VALVE_FAULT.XV05_FAIL_TO_CLOSE,
                      status => "Valves Data".R6_XV05.STATUS);
   END_IF;
END_REGION

REGION Network 61: R6_XV06
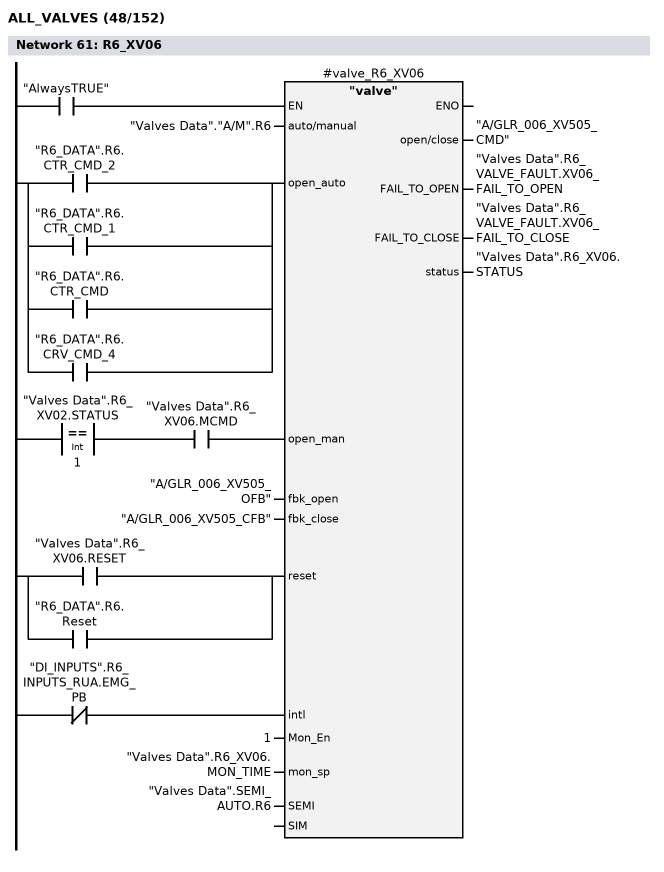
   RUNG wire#powerrail
      Contact( "AlwaysTRUE" )
      #valve_R6_XV06(open_auto := wire#w1, open_man := wire#w2, reset := wire#w3, intl := wire#w4, "auto/manual" := "Valves Data"."A/M".R6, fbk_open := "A/GLR_006_XV505_OFB", fbk_close := "A/GLR_006_XV505_CFB", Mon_En := 1, mon_sp := "Valves Data".R6_XV06.MON_TIME, SEMI := "Valves Data".SEMI_AUTO.R6, SIM :=, "open/close" => "A/GLR_006_XV505_CMD", FAIL_TO_OPEN => "Valves Data".R6_VALVE_FAULT.XV06_FAIL_TO_OPEN, FAIL_TO_CLOSE => "Valves Data".R6_VALVE_FAULT.XV06_FAIL_TO_CLOSE, status => "Valves Data".R6_XV06.STATUS)
   END_RUNG
   RUNG wire#powerrail
      Contact( "R6_DATA".R6.CTR_CMD_2 )
   END_RUNG wire#w1
   RUNG wire#powerrail
      Contact( "R6_DATA".R6.CTR_CMD_1 )
   END_RUNG wire#w1
   RUNG wire#powerrail
      Contact( "R6_DATA".R6.CTR_CMD )
   END_RUNG wire#w1
   RUNG wire#powerrail
      Contact( "R6_DATA".R6.CRV_CMD_4 )
   END_RUNG wire#w1
   RUNG wire#powerrail
      { S7_Templates := "SrcType := Int" } EQ_Contact(in1 := "Valves Data".R6_XV02.STATUS, in2 := 1)
      Contact( "Valves Data".R6_XV06.MCMD )
   END_RUNG wire#w2
   RUNG wire#powerrail
      Contact( "Valves Data".R6_XV06.RESET )
   END_RUNG wire#w3
   RUNG wire#powerrail
      Contact( "R6_DATA".R6.Reset )
   END_RUNG wire#w3
   RUNG wire#powerrail
      I_Contact( "DI_INPUTS".R6_INPUTS_RUA.EMG_PB )
   END_RUNG wire#w4
   // the same network as SCL:
   IF "AlwaysTRUE" THEN
       #valve_R6_XV06("auto/manual" := "Valves Data"."A/M".R6,   // "valve"
                      open_auto := "R6_DATA".R6.CTR_CMD_2 OR "R6_DATA".R6.CTR_CMD_1 OR "R6_DATA".R6.CTR_CMD OR "R6_DATA".R6.CRV_CMD_4,
                      open_man := ("Valves Data".R6_XV02.STATUS = 1) AND "Valves Data".R6_XV06.MCMD,
                      fbk_open := "A/GLR_006_XV505_OFB",
                      fbk_close := "A/GLR_006_XV505_CFB",
                      reset := "Valves Data".R6_XV06.RESET OR "R6_DATA".R6.Reset,
                      intl := NOT "DI_INPUTS".R6_INPUTS_RUA.EMG_PB,
                      Mon_En := 1,
                      mon_sp := "Valves Data".R6_XV06.MON_TIME,
                      SEMI := "Valves Data".SEMI_AUTO.R6,
                      "open/close" => "A/GLR_006_XV505_CMD",
                      FAIL_TO_OPEN => "Valves Data".R6_VALVE_FAULT.XV06_FAIL_TO_OPEN,
                      FAIL_TO_CLOSE => "Valves Data".R6_VALVE_FAULT.XV06_FAIL_TO_CLOSE,
                      status => "Valves Data".R6_XV06.STATUS);
   END_IF;
END_REGION

REGION Network 62: R6_XV07
